(* IEC 61131-3 sources: daoli-st-library/DL_MathData (part 9) *)

(* ---- FC_DL_BcdAddByte.st ---- *)
(*==============================================================================
 * 组件名称 : FC_DL_BcdAddByte ｜ 子库 : DL_MathData ｜ v1.0.0 ｜ 2026-11-23
 * 平台     : CODESYS 3.5 / TwinCAT 3 / InoProShop / Machine Expert（纯 IEC，无厂商库）
 * 功能简介 : 两位 BCD 字节加法：先解码为二进制求和，和 > 99 置错并饱和
 *            到 99，再编码回 BCD。输入含非法 BCD 半字节时置错并返 0。
 * 契约     : 返回 BCD 和 [两位 BCD 形]；xError = TRUE 表示溢出 / 非法输入，
 *            此时返回 99（溢出饱和）或 0（非法输入）；纯函数无状态。
 * 依赖     : 无 DL_ 内部依赖（本批自足实现，不引用库内其他件）
 * 红线自检 : R1 零全局 R2 零%I/%Q R3 纯IEC（*_TO_* 显式转换）
 *            R4 非法 BCD 拒收 + 溢出饱和不回绕 R5 双语注释
 *            R6 N/A（无状态机） R7 N/A（无定时器实例）
 * 修订历史 : 2026-11-23 R78-B1 BCD 校验与算术族模板派生首版
 *============================================================================*)
FUNCTION FC_DL_BcdAddByte : BYTE
VAR_INPUT
    byA : BYTE;         // BCD 加数 / First BCD addend
    byB : BYTE;         // BCD 被加数 / Second BCD addend
END_VAR
VAR_OUTPUT
    xError : BOOL;      // 置错标志：输入非法或和溢出 / Error flag: invalid input or overflow
END_VAR
VAR
    nA : INT;           // byA 解码二进制值 [0..99] / Binary value decoded from byA
    nB : INT;           // byB 解码二进制值 [0..99] / Binary value decoded from byB
    nS : INT;           // 二进制和 [0..99] / Binary sum
    nTens : INT;        // 十位数字 [0..9] / Tens digit
    nOnes : INT;        // 个位数字 [0..9] / Ones digit
END_VAR
xError := FALSE;                    // 置错标志预清 / Preset error flag cleared
FC_DL_BcdAddByte := 16#00;          // 返回值预置 0 / Preset return 0
IF ((byA AND 16#0F) > 16#09) OR (SHR(byA, 4) > 16#09)
    OR ((byB AND 16#0F) > 16#09) OR (SHR(byB, 4) > 16#09) THEN
    xError := TRUE;                 // 输入含非法 BCD 半字节 / Invalid BCD nibble in input
    RETURN;
END_IF
nA := BYTE_TO_INT(SHR(byA, 4)) * 10 + BYTE_TO_INT(byA AND 16#0F);   // 解码 byA / Decode byA
nB := BYTE_TO_INT(SHR(byB, 4)) * 10 + BYTE_TO_INT(byB AND 16#0F);   // 解码 byB / Decode byB
nS := nA + nB;                      // 二进制求和 / Binary sum
IF nS > 99 THEN
    xError := TRUE;                 // 和溢出两位 BCD 域 / Sum overflows two-digit BCD
    nS := 99;                       // 饱和到 99，不回绕 / Saturate at 99, no wrap
END_IF
nTens := nS / 10;                   // 取十位 / Extract tens digit
nOnes := nS MOD 10;                 // 取个位 / Extract ones digit
FC_DL_BcdAddByte := SHL(INT_TO_BYTE(nTens), 4) OR INT_TO_BYTE(nOnes);   // 编码回 BCD / Encode back to BCD
END_FUNCTION

(* ---- FC_DL_BcdDecrementByte.st ---- *)
(*==============================================================================
 * 组件名称 : FC_DL_BcdDecrementByte ｜ 子库 : DL_MathData ｜ v1.0.0 ｜ 2026-11-23
 * 平台     : CODESYS 3.5 / TwinCAT 3 / InoProShop / Machine Expert（纯 IEC，无厂商库）
 * 功能简介 : BCD 字节减 1（如计数值递减）：0 借位回 99（循环计数口径）。
 *            输入含非法 BCD 半字节时防御性返回 0。
 * 契约     : 返回 BCD 减 1 结果 [两位 BCD 形]；非法输入返回 0；
 *            纯函数无状态、同输入同输出。
 * 依赖     : 无 DL_ 内部依赖（本批自足实现，不引用库内其他件）
 * 红线自检 : R1 零全局 R2 零%I/%Q R3 纯IEC（*_TO_* 显式转换）
 *            R4 非法 BCD 返 0 + 0 借位回 99 不越域 R5 双语注释
 *            R6 N/A（无状态机） R7 N/A（无定时器实例）
 * 修订历史 : 2026-11-23 R78-B1 BCD 校验与算术族模板派生首版
 *============================================================================*)
FUNCTION FC_DL_BcdDecrementByte : BYTE
VAR_INPUT
    byVal : BYTE;       // 待递减 BCD 字节 / BCD byte to be decremented
END_VAR
VAR
    nV : INT;           // 解码二进制值 [0..99] / Decoded binary value
    nTens : INT;        // 十位数字 [0..9] / Tens digit
    nOnes : INT;        // 个位数字 [0..9] / Ones digit
END_VAR
FC_DL_BcdDecrementByte := 16#00;    // 返回值预置 0 / Preset return 0
IF ((byVal AND 16#0F) > 16#09) OR (SHR(byVal, 4) > 16#09) THEN
    RETURN;                         // 非法 BCD 输入防御性返 0 / Invalid BCD input returns 0
END_IF
nV := BYTE_TO_INT(SHR(byVal, 4)) * 10 + BYTE_TO_INT(byVal AND 16#0F);   // 解码 / Decode
nV := nV - 1;                       // 二进制减 1 / Decrement in binary
IF nV < 0 THEN
    nV := 99;                       // 0 借位回 99 / Borrow 0 back to 99
END_IF
nTens := nV / 10;                   // 取十位 / Extract tens digit
nOnes := nV MOD 10;                 // 取个位 / Extract ones digit
FC_DL_BcdDecrementByte := SHL(INT_TO_BYTE(nTens), 4) OR INT_TO_BYTE(nOnes);     // 编码回 BCD / Encode back to BCD
END_FUNCTION

(* ---- FC_DL_BcdIncrementByte.st ---- *)
(*==============================================================================
 * 组件名称 : FC_DL_BcdIncrementByte ｜ 子库 : DL_MathData ｜ v1.0.0 ｜ 2026-11-23
 * 平台     : CODESYS 3.5 / TwinCAT 3 / InoProShop / Machine Expert（纯 IEC，无厂商库）
 * 功能简介 : BCD 字节加 1（如计数器 / 计数值递增）：99 进位回 0。
 *            输入含非法 BCD 半字节时防御性返回 0。
 * 契约     : 返回 BCD 加 1 结果 [两位 BCD 形]；非法输入返回 0；
 *            纯函数无状态、同输入同输出。
 * 依赖     : 无 DL_ 内部依赖（本批自足实现，不引用库内其他件）
 * 红线自检 : R1 零全局 R2 零%I/%Q R3 纯IEC（*_TO_* 显式转换）
 *            R4 非法 BCD 返 0 + 99 进位回 0 不越域 R5 双语注释
 *            R6 N/A（无状态机） R7 N/A（无定时器实例）
 * 修订历史 : 2026-11-23 R78-B1 BCD 校验与算术族模板派生首版
 *============================================================================*)
FUNCTION FC_DL_BcdIncrementByte : BYTE
VAR_INPUT
    byVal : BYTE;       // 待递增 BCD 字节 / BCD byte to be incremented
END_VAR
VAR
    nV : INT;           // 解码二进制值 [0..99] / Decoded binary value
    nTens : INT;        // 十位数字 [0..9] / Tens digit
    nOnes : INT;        // 个位数字 [0..9] / Ones digit
END_VAR
FC_DL_BcdIncrementByte := 16#00;    // 返回值预置 0 / Preset return 0
IF ((byVal AND 16#0F) > 16#09) OR (SHR(byVal, 4) > 16#09) THEN
    RETURN;                         // 非法 BCD 输入防御性返 0 / Invalid BCD input returns 0
END_IF
nV := BYTE_TO_INT(SHR(byVal, 4)) * 10 + BYTE_TO_INT(byVal AND 16#0F);   // 解码 / Decode
nV := nV + 1;                       // 二进制加 1 / Increment in binary
IF nV > 99 THEN
    nV := 0;                        // 99 进位回 0 / Carry 99 back to 0
END_IF
nTens := nV / 10;                   // 取十位 / Extract tens digit
nOnes := nV MOD 10;                 // 取个位 / Extract ones digit
FC_DL_BcdIncrementByte := SHL(INT_TO_BYTE(nTens), 4) OR INT_TO_BYTE(nOnes);     // 编码回 BCD / Encode back to BCD
END_FUNCTION

(* ---- FC_DL_BcdIsValidByte.st ---- *)
(*==============================================================================
 * 组件名称 : FC_DL_BcdIsValidByte ｜ 子库 : DL_MathData ｜ v1.0.0 ｜ 2026-11-23
 * 平台     : CODESYS 3.5 / TwinCAT 3 / InoProShop / Machine Expert（纯 IEC，无厂商库）
 * 功能简介 : 判定字节是否为合法两位 BCD 编码：高 / 低半字节均须 <= 9
 *            （0x0A..0x0F 非法）。纯位运算实现，不用库函数。
 * 契约     : 返回 TRUE = 合法 BCD 字节（00..99 的 BCD 形）；输入 byVal
 *            任意字节；纯函数无状态、同输入同输出。
 * 依赖     : 无 DL_ 内部依赖（本批自足实现）
 * 红线自检 : R1 零全局 R2 零%I/%Q R3 纯IEC R4 半字节越 9 拒收
 *            R5 双语注释 R6 N/A（无状态机） R7 N/A（无定时器实例）
 * 修订历史 : 2026-11-23 R78-B1 BCD 校验与算术族模板派生首版
 *============================================================================*)
FUNCTION FC_DL_BcdIsValidByte : BOOL
VAR_INPUT
    byVal : BYTE;       // 待判定字节 / Byte to be validated
END_VAR
IF ((byVal AND 16#0F) > 16#09) OR (SHR(byVal, 4) > 16#09) THEN
    FC_DL_BcdIsValidByte := FALSE;      // 任一半字节 > 9：非法 BCD / Any nibble > 9: invalid BCD
ELSE
    FC_DL_BcdIsValidByte := TRUE;       // 高低半字节均 <= 9：合法 / Both nibbles <= 9: valid
END_IF
END_FUNCTION

(* ---- FC_DL_BcdIsValidWord.st ---- *)
(*==============================================================================
 * 组件名称 : FC_DL_BcdIsValidWord ｜ 子库 : DL_MathData ｜ v1.0.0 ｜ 2026-11-23
 * 平台     : CODESYS 3.5 / TwinCAT 3 / InoProShop / Machine Expert（纯 IEC，无厂商库）
 * 功能简介 : 判定 16 位字是否为合法 4 位 BCD 编码：4 个半字节均须 <= 9
 *            （任一半字节 0x0A..0x0F 非法）。纯位运算 FOR 循环实现，
 *            不用库函数。
 * 契约     : 返回 TRUE = 合法 BCD 字（0000..9999 的 BCD 形）；输入 wVal
 *            任意字；循环轮次固定 4，结构有界；纯函数无状态。
 * 依赖     : 无 DL_ 内部依赖（本批自足实现）
 * 红线自检 : R1 零全局 R2 零%I/%Q R3 纯IEC R4 半字节越 9 拒收 + FOR 上界常量
 *            R5 双语注释 R6 N/A（无状态机） R7 N/A（无定时器实例）
 * 修订历史 : 2026-11-23 R78-B1 BCD 校验与算术族模板派生首版
 *============================================================================*)
FUNCTION FC_DL_BcdIsValidWord : BOOL
VAR_INPUT
    wVal : WORD;        // 待判定 16 位字 / Word to be validated
END_VAR
VAR
    i : INT;            // 半字节序号 0..3 / Nibble index 0..3
END_VAR
FC_DL_BcdIsValidWord := TRUE;       // 预置合法，逐位复核 / Preset valid, recheck nibble by nibble
FOR i := 0 TO 3 DO                  // 4 个半字节逐一校验 / Check all 4 nibbles
    IF (SHR(wVal, i * 4) AND 16#000F) > 16#0009 THEN
        FC_DL_BcdIsValidWord := FALSE;      // 该半字节 > 9：非法 BCD / Nibble > 9: invalid BCD
    END_IF
END_FOR
END_FUNCTION

(* ---- FC_DL_BcdSubByte.st ---- *)
(*==============================================================================
 * 组件名称 : FC_DL_BcdSubByte ｜ 子库 : DL_MathData ｜ v1.0.0 ｜ 2026-11-23
 * 平台     : CODESYS 3.5 / TwinCAT 3 / InoProShop / Machine Expert（纯 IEC，无厂商库）
 * 功能简介 : 两位 BCD 字节减法：先解码为二进制求差，差 < 0（借位下溢）
 *            置错并饱和到 0，再编码回 BCD。输入含非法 BCD 半字节时置错
 *            并返 0。
 * 契约     : 返回 BCD 差 [两位 BCD 形]；xError = TRUE 表示下溢 / 非法输入，
 *            此时返回 0（下溢饱和）；纯函数无状态。
 * 依赖     : 无 DL_ 内部依赖（本批自足实现，不引用库内其他件）
 * 红线自检 : R1 零全局 R2 零%I/%Q R3 纯IEC（*_TO_* 显式转换）
 *            R4 非法 BCD 拒收 + 下溢饱和不回绕 R5 双语注释
 *            R6 N/A（无状态机） R7 N/A（无定时器实例）
 * 修订历史 : 2026-11-23 R78-B1 BCD 校验与算术族模板派生首版
 *============================================================================*)
FUNCTION FC_DL_BcdSubByte : BYTE
VAR_INPUT
    byA : BYTE;         // BCD 被减数 / BCD minuend
    byB : BYTE;         // BCD 减数 / BCD subtrahend
END_VAR
VAR_OUTPUT
    xError : BOOL;      // 置错标志：输入非法或借位下溢 / Error flag: invalid input or borrow underflow
END_VAR
VAR
    nA : INT;           // byA 解码二进制值 [0..99] / Binary value decoded from byA
    nB : INT;           // byB 解码二进制值 [0..99] / Binary value decoded from byB
    nD : INT;           // 二进制差 [0..99] / Binary difference
    nTens : INT;        // 十位数字 [0..9] / Tens digit
    nOnes : INT;        // 个位数字 [0..9] / Ones digit
END_VAR
xError := FALSE;                    // 置错标志预清 / Preset error flag cleared
FC_DL_BcdSubByte := 16#00;          // 返回值预置 0 / Preset return 0
IF ((byA AND 16#0F) > 16#09) OR (SHR(byA, 4) > 16#09)
    OR ((byB AND 16#0F) > 16#09) OR (SHR(byB, 4) > 16#09) THEN
    xError := TRUE;                 // 输入含非法 BCD 半字节 / Invalid BCD nibble in input
    RETURN;
END_IF
nA := BYTE_TO_INT(SHR(byA, 4)) * 10 + BYTE_TO_INT(byA AND 16#0F);   // 解码 byA / Decode byA
nB := BYTE_TO_INT(SHR(byB, 4)) * 10 + BYTE_TO_INT(byB AND 16#0F);   // 解码 byB / Decode byB
nD := nA - nB;                      // 二进制求差 / Binary difference
IF nD < 0 THEN
    xError := TRUE;                 // 借位下溢出两位 BCD 域 / Borrow underflow
    nD := 0;                        // 饱和到 0，不回绕 / Saturate at 0, no wrap
END_IF
nTens := nD / 10;                   // 取十位 / Extract tens digit
nOnes := nD MOD 10;                 // 取个位 / Extract ones digit
FC_DL_BcdSubByte := SHL(INT_TO_BYTE(nTens), 4) OR INT_TO_BYTE(nOnes);   // 编码回 BCD / Encode back to BCD
END_FUNCTION

(* ---- FC_DL_BcdToByte.st ---- *)
(*
    FC_DL_BcdToByte —— 2 位半字节 BCD 解码（BYTE 容器）
    ------------------------------------------------------------------
    分类      : DL_MathData / Convert
    前缀      : FC_DL_
    版本      : 1.0.0
    溯源      : IEC 61131-3 标准语义的道莅防御性实现（BYTE 容器 2 位 BCD → USINT 数值）；
                域内委托平台内建 BCD_TO_BYTE，本件不重实现数学内核；
                半字节合法性校验、满量程提示、错误分级与码位 100% 自有；
                clean-room 重写，未复制任何闭源厂商源码，参考实现仅限 MIT/Apache 许可
    平台      : 纯 IEC 61131-3，CODESYS V3.5+ / TwinCAT 3 / InoProShop 通用
    作者      : 道莅代码库 · PLC编程专家（R20）
    ------------------------------------------------------------------
    功能说明  : 拨码开关组态位、老式仪表组态字最常见的 2 位 BCD 编码（一个 BYTE 装 0~99），
                解码成 0~99 的数值参与比对。
                核心防御：① 先判后算——两个半字节都必须 ≤ 9 才允许进内建。
                   非法 BCD（如 16#1F、16#AA）在内建层的行为平台各不相同（有的翻转、
                   有的返回原值、有的置 0），是本件最不能容忍的不确定点；
                ② 校验只看半字节数值，不看容器大小，故 16#99 合法、16#FF 非法；
                ③ 满量程 99 发信息级提示：拨码全拨到 9 常是调试残留，
                   值本身合法，不该升故障级；
                ④ 合成路径（若平台缺内建）在容器校验之后做半字节乘加，
                   属校验后合成，不是重实现数学内核。
                职责边界：反向编码归 FC_DL_ByteToBcd；4 位 Word 容器归 FC_DL_BcdToWord，
                8 位 Udint 容器归 FC_DL_BcdToUdint；本件只管 2 位拨码容器。
    编译门槛  : 主路径依赖平台内建 BCD_TO_BYTE，三平台标准库均提供。
                若目标平台缺该内建，按合成路径落地：uOut = uHi * 10 + uLo，
                两半字节已由段 2 保证 ≤ 9，乘加结果必然 ≤ 99，无溢出可能。
    错误码    : 16#0001_041C BCD 值恰为满量程 99（多拨码开关调试残留）——信息级，值可用
                16#0001_041D 预留禁用（信息级，不得挪用）
                16#0001_0348 非法 BCD（某半字节 > 9）——故障级，返回 0
                16#0001_0349 预留（故障级，不得挪用）
                16#0001_034A 预留禁用（故障级，不得挪用）
    码位总账  : 16#0001_041C 用 / 16#0001_041D 预留 ｜ 16#0001_0348 用 / 16#0001_0349 预留 / 16#0001_034A 预留
    状态机    : R6 标注 N/A —— 本组件为纯函数无顺序状态机，无 CASE 可写，非法状态不可能出现
    采样约定  : 本件无定时器、无沿检测、无状态；单拍纯计算，结论与任务周期无关。
    修订记录  : 2026-11-16 v1.0.0 首次入库（R20）
*)
FUNCTION FC_DL_BcdToByte : USINT
VAR_INPUT
    uBcd             : BYTE;                  // BCD 编码值 [无量纲]，每半字节 0~9，合计 0~99 / BCD value [dimensionless], each nibble 0 to 9, total 0 to 99
END_VAR
VAR_OUTPUT
    eErr             : UDINT;                 // 错误码，0=正常 / error id, 0=ok
    bError           : BOOL;                  // 故障标志，eErr 为故障级时 TRUE / error flag, TRUE on fault-level eErr
    bValid           : BOOL;                  // 返回值是否可用（非法 BCD 为 FALSE）/ return usable, FALSE on an illegal BCD
END_VAR
VAR CONSTANT
    DL_BCD_NIB_MAX   : BYTE := 9;             // 单个半字节的合法上限 [无量纲] / legal upper bound of one nibble [dimensionless]
    DL_BCD_MASK_LO   : BYTE := 16#0F;         // 低半字节掩码 [位图] / low nibble mask [bitmap]
    DL_BCD_SHIFT_HI  : USINT := 4;            // 高半字节移位量 [bit]，结构性小于 8 / the high nibble shift [bit], structurally below 8
    DL_BCD_FULL      : USINT := 99;           // 满量程值，用于提示 [无量纲] / full scale value used by the hint [dimensionless]
    DL_USINT_ZERO    : USINT := 0;            // 无符号零常量，避免裸字面量 [无量纲] / unsigned zero constant [dimensionless]
END_VAR
VAR
    uLo              : BYTE;                  // 低半字节 [无量纲] / the low nibble [dimensionless]
    uHi              : BYTE;                  // 高半字节 [无量纲] / the high nibble [dimensionless]
    uOut             : USINT;                 // 结果中间量 [无量纲] / result intermediate [dimensionless]
END_VAR

// 段 1｜返回值与错误状态预置 / segment 1, preset return value and error status
FC_DL_BcdToByte := DL_USINT_ZERO;             // 故障缺省返回 0 [无量纲] / fault default returns zero [dimensionless]
eErr := 0;                                    // 预置无错误 / preset no error
bError := FALSE;                              // 预置无故障 / preset no fault
bValid := FALSE;                              // 预置不可用，通过闸门后置位 / preset invalid, set TRUE after the gates
uOut := DL_USINT_ZERO;                        // 结果中间量清零 / clear the result intermediate

// 段 2｜半字节分解与合法性校验（先判后算，域外绝不进内建）/ segment 2, nibble split and legality gate
uLo := uBcd AND DL_BCD_MASK_LO;               // 低半字节 [无量纲] / extract the low nibble [dimensionless]
uHi := SHR(uBcd, DL_BCD_SHIFT_HI);            // 高半字节，移位量 4 结构性小于 8 [无量纲] / extract the high nibble, the shift stays below 8 [dimensionless]

IF (uLo > DL_BCD_NIB_MAX) OR (uHi > DL_BCD_NIB_MAX) THEN
    eErr := 16#0001_0348;                     // 故障级：非法 BCD，半字节超 9 / fault level, illegal BCD, a nibble exceeds nine
    bError := TRUE;                           // 置故障标志 / raise the error flag
    bValid := FALSE;                          // 返回值不可用 / flag the return as unusable
    FC_DL_BcdToByte := DL_USINT_ZERO;         // 确定缺省值 0 / deterministic default of zero
    RETURN;                                   // 出口，不触碰内建 / exit, the built-in is never touched
END_IF

// 段 3｜主体：容器校验通过后委托平台内建 / segment 3, delegate the built-in after the container check
uOut := BYTE_TO_USINT(BCD_TO_BYTE(uBcd));     // BCD → 数值 [无量纲] / decode BCD into a number [dimensionless]

// 段 4｜发布结果与满量程提示（信息级，不置 bError）/ segment 4, publish and hint the full scale value
FC_DL_BcdToByte := uOut;                      // 输出解码值 0~99 [无量纲] / publish the decoded value 0 to 99 [dimensionless]
bValid := TRUE;                               // 合法 BCD 即可用 / a legal BCD is usable
IF uOut = DL_BCD_FULL THEN
    eErr := 16#0001_041C;                     // 信息级：满量程 99，多为拨码调试残留 / info level, full scale, often left over from commissioning
END_IF
END_FUNCTION

(* ---- FC_DL_BcdToDint.st ---- *)
(*
  ==================================================================
  组件名 Component  : FC_DL_BcdToDint
  分类   Category   : DL_MathData
  前缀   Naming     : FC_DL_ ｜ b/n/u/f/t/e/st 类型前缀制（R265）
  码位   Code ID    : 16#0001_0657（故障级）
  版本   Version    : 1.0.0
  复杂度 Complexity  : 低
  功能   Purpose    : 8 位 BCD（DWORD 容器，8 个半字节）→ DINT，逐码元合法性闸，
                      任一半字节 > 9 判故障早退，禁静默按半字节折算。
  开源溯源 Origin    : 公开公式 clean-room，参考 BCD 编码公开工程语义（分类与参数域
                      借鉴，零代码复制），本件实现、闸门与码位 100% 自有。
  许可证 License    : MIT
  参考   Reference  : IEC 61131-3:2013 §6.6 移位与位运算符（SHR / AND）
  平台   Platform   : 纯 IEC 61131-3（FOR / SHR / AND / 四则），三平台通用
  依赖   Depends    : 仅 Standard.library（无库调用）
  分工声明 Split     : FC_DL_BcdToByte / FC_DL_BcdToWord / FC_DL_BcdToUdint 为既有
                      BCD 解码族（BYTE / WORD / UDINT 位宽），本件补 DWORD 8 位宽
                      解码口，四件互引（R216）。
  归属 Ownership     : 本件无 TYPE 声明；全部引脚为 IEC 标准原生类型。
  ------------------------------------------------------------------
  边界 Boundary     :
                      一 域证明（写死）：8 位 BCD 最大 99999999 < 2147483647（DINT
                         上界），累加无溢出可能，故本件无溢出分支；
                      二 逐码元提取：SHR 移位量 4·k（k = 0..7）最大 28 < 32（DWORD
                         位宽），结构性安全（R48 移位量归一：移位量上界由循环界
                         常量证明，禁运行时可变移位量越位宽）；
                      三 任一码元 > 9 → 故障级码 + bBadDigit = TRUE + nOut = 0 +
                         三件套 + RETURN 早退（禁把 A~F 半字节静默折算）；
                      四 首个非法码元即早退（首因保序），bBadDigit 单点置位；
                      五 纯函数：无记忆量、无定时器、无边沿实例，每调用重算；
                      六 无全局、无外部变量、无物理地址、无指针。
  错误码 Codes      :
    16#0001_0657【故障级】非法码元（8 个半字节任一 > 9，首个非法位即早退）
  码位反证 Note     :
    本件仅一个故障场景：8 个码元的合法性出口组合完全同形（nOut = 0、bBadDigit =
    TRUE、bValid = FALSE），无法从输出区分「哪一位非法」，按 R90 只立一码，
    非法位序号不外显（如需位级定位由调用方自行逐半字节复扫）。
  验收 Acceptance   :
    算法已证（脚本）：未跑 ｜ 编译器已证（三平台）：未跑
    V1 16#00000000 → 0；V2 16#99999999 → 99999999（精确无溢出）
    V3 16#0000000A → 故障 0657 + bBadDigit（禁折算）
    V4 16#12345678 → 12345678；V5 16#00000007 → 7（前导零）
    V6 高位半字节 16#A0000000 与低位 16#0000000F → 均故障（A/F 两端抽验）
  修订记录 Revision  :
    2026-11-21  v1.0.0  R63 首版（批 1 · 序号 1）
  ==================================================================
*)
FUNCTION FC_DL_BcdToDint : BOOL
VAR_INPUT
    udBcd   : DWORD := 16#00000000; // 8 位 BCD 输入 [码]，8 个半字节 / the eight digit BCD input in a double word container
END_VAR
VAR_OUTPUT
    nOut    : DINT := 0;            // 解码结果 [个]，非法码元时为 0 / the decoded result, zero when a digit is illegal
    bBadDigit : BOOL := FALSE;      // 非法码元标志（任一半字节 > 9）[-] / the illegal digit flag raised when any nibble exceeds nine
    bValid  : BOOL := FALSE;        // 结果可用 [-] / the result usable flag
    eErr    : UDINT := 16#0000_0000; // 错误码，0 = 正常 / the error code, zero is ok
    bError  : BOOL := FALSE;        // 故障标志（故障级码同拍置位，R45 配对）/ the fault flag raised with a fault level code
END_VAR
VAR
    k       : DINT := 0;  // 半字节遍历索引 [下标]，0..7 / the nibble traversal index from zero to seven
    nShift  : DINT := 0;  // 移位量 [位]，4·k ≤ 28 结构性安全 / the shift amount of four times the index, proven below the word width
    uDig    : USINT := 0; // 当前半字节码元 [位] / the current digit nibble
    nAcc    : DINT := 0;  // 十进制累加器（Horner 展开）[个] / the decimal accumulator of the Horner expansion
END_VAR  // R64 结构补齐：VAR 段缺失的 END_VAR（门禁机械修复）
VAR CONSTANT
    DL_BCD_MASK  : DWORD := 16#0000000F; // 半字节掩码常量（提级禁魔法数）[-] / the nibble mask constant lifted out of the body
    DL_BCD_DIG9  : USINT := 9;           // 合法码元上界 [位] / the legal digit ceiling of nine
    DL_BCD_NIB   : DINT := 4;            // 每码元位宽 [位] / the nibble width of four bits
    DL_BCD_N     : DINT := 8;            // 码元总数 [个]（DWORD 恰 8 半字节，R57）/ the nibble count of eight aligned with the container
    DL_BCD_ZERO  : DINT := 0;            // 整型零常量 [个] / the integer zero constant
    DL_BCD_ONE   : DINT := 1;            // 整型一常量 [个] / the integer one constant
    DL_BCD_TEN   : DINT := 10;           // 十进制权值基数 [个] / the decimal weight base of ten
END_VAR

// 段 1｜返回值与全部出口预置安全值（R45 四段式第一段）/ segment 1, the preset of the return and every outlet
FC_DL_BcdToDint := FALSE; // 返回值预置假 / preset the return false
nOut := DL_BCD_ZERO; // 结果预置零 [个] / preset the result zero
bBadDigit := FALSE; // 非法码元标志预置假 / preset the illegal digit flag false
bValid := FALSE; // 可用标志预置假 / preset the validity false
eErr := 16#0000_0000; // 错误码预置正常 / preset the code to ok
bError := FALSE; // 故障标志预置假 / preset the error flag false
nAcc := DL_BCD_ZERO; // 累加器预置零 [个] / preset the accumulator zero
k := DL_BCD_ZERO; // 索引预置零 / preset the index zero
nShift := DL_BCD_ZERO; // 移位量预置零 [位] / preset the shift amount zero
uDig := 0; // 码元预置零 [位] / preset the digit zero

// 段 2｜逐码元提取与合法性闸（移位量 4·k ≤ 28 < 32 结构性安全，边界二）/ segment 2, the digit extraction with the structural shift bound
FOR k := DL_BCD_ZERO TO DL_BCD_N - DL_BCD_ONE DO // 有界遍历 8 个半字节（循环界常量证明，无死循环）/ the bounded traversal over eight nibbles proven by the constant loop bound
    nShift := DL_BCD_NIB * k; // 移位量 = 4·k，最大 28 [位] / the shift amount of four times the index, at most twenty eight
    uDig := DWORD_TO_USINT(SHR(udBcd, nShift) AND DL_BCD_MASK); // 提取当前半字节（SHR 后与掩码，常量提级）/ extract the current nibble by shifting then masking with the lifted constant
    IF uDig > DL_BCD_DIG9 THEN // 码元 > 9：非法（边界三，禁折算）/ a digit above nine is illegal, never folded silently
        bBadDigit := TRUE; // 置非法码元标志 / raise the illegal digit flag
        eErr := 16#0001_0657; // 故障级：非法码元 / fault grade, an illegal digit
        bError := TRUE; // 同拍置故障标志（R45 配对）/ raise the fault flag on the same scan
        bValid := FALSE; // 结果不可用 / the result is not usable
        nOut := DL_BCD_ZERO; // 结果强制归零（禁部分折算值外泄）/ force the result to zero so no partial fold leaks
        RETURN; // 早退（首因保序，边界四）/ early return with the first cause kept
    END_IF
    nAcc := (nAcc * DL_BCD_TEN) + USINT_TO_DINT(uDig); // Horner 十进制累加：nAcc = nAcc×10 + 码元 [个] / the Horner decimal accumulation, the domain proof in boundary one covers every step
END_FOR

// 段 3｜统一出口（域证明：nAcc ≤ 99999999 < DINT 上界，无溢出分支，边界一）/ segment 3, the unified outlet with the domain proof
nOut := nAcc; // 结果出口 [个] / the result outlet
bValid := TRUE; // 结果可用 / the result is usable
FC_DL_BcdToDint := TRUE; // 返回成功 / return success
END_FUNCTION

(* ---- FC_DL_BcdToUdint.st ---- *)
(*
    FC_DL_BcdToUdint —— 8 位十进制 BCD 码到 UDINT 防御转换
    ------------------------------------------------------------------
    分类      : DL_MathData / Convert
    前缀      : FC_DL_
    版本      : 1.0.0
    溯源      : IEC 61131-3 标准语义的道莅防御性实现
                （内部委托平台内建函数，外围统一错误码/钳位/双语文档；
                  未复制任何闭源厂商源码，参考实现仅限 MIT/Apache 许可）
    平台      : 纯 IEC 61131-3，CODESYS / TwinCAT / InoProShop 通用
    作者      : 道莅代码库 · PLC编程专家（R16）
    ------------------------------------------------------------------
    功能说明  : 将 8 位十进制 BCD 码输入（每半字节 0~9）防御性转换为 UDINT 并返回；
                逐半字节合法性校验：任一半字节值 > 9（即 16#A~16#F 非法 BCD 码）判为
                故障级 16#0001_02A6，返回 0 且 bValid=FALSE；
                域内按半字节以 10 为基加权累加还原十进制值（乘子为常量基 10 的幂，
                最大权值 10^7、最大累加和 99999999，均在 UDINT 域内无溢出）；
                校验覆盖范围说明：UDINT 为 32 位容器，恰含 8 个 BCD 半字节（k=0..7），
                完整覆盖 8 位十进制域 0..99999999；k=8..15 的半字节在 32 位容器中不存在，
                且移位量 ≥32 属跨平台未定义行为，故不实施越界校验；
                本组件无钳位路径（非法半字节直接故障拦截，域内值精确还原）。
    错误码    : 16#0001_02A6 存在非法 BCD 半字节（半字节值 16#A~16#F）——故障级，返回 0
                16#0001_01D0 预留禁用（信息级，不得挪用）
                16#0001_01D1 预留禁用（信息级，不得挪用）
                16#0001_02A7 预留禁用（故障级，不得挪用）
                16#0001_02A8 预留禁用（故障级，不得挪用）
    状态机    : R6 标注 N/A —— 本组件为纯函数无顺序状态机，无 CASE 可写，非法状态不可能出现，故以本节说明替代 ELSE 兜底
    修订记录  : 2026-11-16 v1.0.0 首次入库（R16）
*)
FUNCTION FC_DL_BcdToUdint : UDINT
VAR_INPUT
    uBcd : UDINT; // 8 位十进制 BCD 码 [BCD 位]，每半字节 0~9 / 8-digit BCD code, each nibble 0~9
END_VAR
VAR_OUTPUT
    eErr   : UDINT; // 错误码，0=正常 / error id, 0=ok
    bError : BOOL;  // 是否出错，eErr 非 0 时为 TRUE / error flag, TRUE when eErr is nonzero
    bValid : BOOL;  // 输出是否有效可用 / output valid flag
END_VAR
VAR CONSTANT
    DL_BCD_NIB_MASK : UDINT := 16#F;  // 半字节掩码 [BCD 位] / nibble mask
    DL_BCD_NIB_MAX  : UDINT := 16#9;  // 合法 BCD 半字节上界 9 [BCD 位] / valid BCD nibble upper bound 9
    DL_BCD_NIB_CNT  : INT   := 8;     // UDINT 32 位容器 BCD 半字节总数 [个] / total BCD nibble count of 32-bit UDINT container
    DL_DEC_BASE     : UDINT := 10;    // 十进制加权基 [基数] / decimal weighting base
END_VAR
VAR
    i       : INT;   // 半字节循环索引 [个] / nibble loop index
    uNib    : UDINT; // 当前半字节值 [BCD 位] / current nibble value
    uWeight : UDINT; // 当前半字节十进制权值（10^i） [倍] / current nibble decimal weight (10^i)
END_VAR

// 段 1｜返回值与错误状态预置 / segment 1, preset return value and error status
FC_DL_BcdToUdint := 0; // 故障缺省返回 0 [无量纲] / fault default returns 0
eErr   := 0;     // 预置无错误 / preset no error
bError := FALSE; // 预置无故障 / preset no fault
bValid := FALSE; // 预置无效，通过全半字节校验后置位 / preset invalid, set TRUE after all-nibble check passes

// 段 2｜逐半字节校验与十进制加权累加（末段） / segment 2, per-nibble validation and decimal weighted accumulation (final)
uWeight := 1; // 最低半字节权值 10^0 [倍] / lowest nibble weight 10^0
FOR i := 0 TO DL_BCD_NIB_CNT - 1 DO
    uNib := SHR(uBcd, 4 * i) AND DL_BCD_NIB_MASK; // 取第 i 个半字节（SHR 移位量 4*i ≤ 28 安全） / extract i-th nibble (shift 4*i <= 28, safe)
    IF uNib > DL_BCD_NIB_MAX THEN
        FC_DL_BcdToUdint := 0;    // 故障级返回 0，清除部分累加值 / fault level returns 0, clear partial accumulation
        eErr   := 16#0001_02A6;   // 非法 BCD 半字节故障码 / invalid BCD nibble fault id
        bError := TRUE;           // 置故障标志 / set fault flag
        bValid := FALSE;          // 输出无效 / output invalid
        RETURN;                   // 立即返回 / immediate return
    END_IF
    FC_DL_BcdToUdint := FC_DL_BcdToUdint + uNib * uWeight; // 半字节加权累加（最大 99999999 无溢出） / weighted accumulation (max 99999999, no overflow)
    uWeight := uWeight * DL_DEC_BASE; // 权值升位 ×10（最大 10^7，UDINT 域内无溢出） / weight times 10 (max 10^7, no UDINT overflow)
END_FOR
bError := FALSE; // 全部半字节合法，无故障 / all nibbles valid, no fault
bValid := TRUE;  // 输出有效可用 / output valid
END_FUNCTION

(* ---- FC_DL_BilinearInterp.st ---- *)
(*
  ==================================================================
  组件名 Component  : FC_DL_BilinearInterp
  分类   Category   : DL_MathData
  版本   Version    : 1.0.0
  功能   Purpose    : 双线性插值：在等距网格表上按 (fX, fY) 求插值。
                      越界策略=「钳位到边界单元并置码不静默」（头注定稿口径）：
                      fX/fY 超出 [fX0, fX0+(n-1)*d] 时钳到边界单元继续插值，
                      输出有效但带码 02；末端格点用 1E-9 容差处理防 i1 越界
                      一行（fU 恰好等于上界时 i0 退到 n-2、tx 收满 1.0，
                      n=1 退化为常量直通）。
  来源   Source     : t2-1-lgf-math（数学族：双线性插值为公开数值方法口径，
                      实现零源码复制）
  互引   Cross-ref  : FC_DL_InterpolateTable3D（同族三维插值原子，本件为其
                      二维退化对偶，可级联使用）
  平台   Platform   : 纯 IEC 61131-3 四则 + TRUNC，三平台通用
  依赖   Depends    : 无 DL_ 内部依赖；无标准库
  表格口径 Table    : aTable 为定长容量数组（NY_MAX × NX_MAX 见常量段），
                      实际使用 ny=nRows / nx=nCols 由输入给定，容量外元素
                      永不访问（下标闸先行）；行序 = [y 索引][x 索引]。
  红线   Redline    : R1 零全局/VAR_EXTERNAL/R2 零 %I/%Q/R3 纯 IEC 标准
                      R4 步距≤0 与行列数<1 配置闸 + 元素级非有限闸（含四角
                      值）+ 越界钳位显式置码 + 除法分母已闸
                      R5 全变量双语同行注释/R6 纯函数无状态机（CASE 不适用）
                      R7 无定时器与沿检测/R8 容差与容量常量化
  错误码 Codes      : 01【失效级】配置非法（nRows/nCols < 1 或步距 ≤ 0 或
                      行列数超容量），返回 0
                      02【信息级】fX/fY 越界已钳位到边界单元（输出有效）
                      03【失效级】任一输入或四角表值非有限，返回 0
  码位反证 Note     : 02 与 03 分立依据（R90）：02 时 bValid=TRUE 带码、
                      03 时 bValid=FALSE，双通道可唯一区分；01 与 03 分立：
                      01 在配置面可观测、03 在数据面可观测，入口不同。
  验收   Acceptance : V1 网格中心点 → 精确双线性值 ｜ V2 fX 超上界 → 钳边界
                      + 码 02 ｜ V3 fDx=0 → 码 01 ｜ V4 nCols=1 → y 向插值
                      常量直通 ｜ V5 表值 NaN → 码 03 ｜ V6 末端格点容差 →
                      不越界不置 02
  变更   Revision   : 2026-11-22  v1.0.0  R66 首版（编码阶段批 2 序 5）
  ==================================================================
*)
FUNCTION FC_DL_BilinearInterp : LREAL
VAR_INPUT
    aTable : ARRAY[0..BIL_NY_MAX - 1, 0..BIL_NX_MAX - 1] OF LREAL; // 容量网格表 [表值]（实际 ny/nx 由 nRows/nCols 给定，行序=[y][x]）/ the capacity grid table
    nRows  : UDINT;  // 实际行数（y 向格点数）[个]，≥1 / the actual rows, at least one
    nCols  : UDINT;  // 实际列数（x 向格点数）[个]，≥1 / the actual columns, at least one
    fX     : LREAL;  // 查询点 x 坐标 [物理单位同表] / the query x coordinate
    fY     : LREAL;  // 查询点 y 坐标 [物理单位同表] / the query y coordinate
    fX0    : LREAL;  // x 起始格点坐标 [物理单位同表] / the x grid origin
    fDx    : LREAL;  // x 步距 [物理单位同表]，须 > 0 / the x step, must be positive
    fY0    : LREAL;  // y 起始格点坐标 [物理单位同表] / the y grid origin
    fDy    : LREAL;  // y 步距 [物理单位同表]，须 > 0 / the y step, must be positive
END_VAR
VAR_OUTPUT
    bValid : BOOL;   // 输出可用标志（码 02 时仍 TRUE）[-] / the output usable flag, true also with code 02
    nErrId : UDINT;  // 错误码，0=正常，01/02/03 见头注 [码] / the error code [code]
END_VAR
VAR
    fU     : LREAL;  // x 向规格化浮点下标 [格] / the normalized floating x index [cell]
    fV     : LREAL;  // y 向规格化浮点下标 [格] / the normalized floating y index [cell]
    fXmax  : LREAL;  // x 上边界格点坐标 [物理单位] / the x upper boundary coordinate
    fYmax  : LREAL;  // y 上边界格点坐标 [物理单位] / the y upper boundary coordinate
    ix0    : UDINT;  // x 向左格点下标 [格] / the left x cell index
    ix1    : UDINT;  // x 向右格点下标 [格] / the right x cell index
    iy0    : UDINT;  // y 向下格点下标 [格] / the lower y cell index
    iy1    : UDINT;  // y 向上格点下标 [格] / the upper y cell index
    fTx    : LREAL;  // x 向格内分数 0~1 [-] / the in cell x fraction
    fTy    : LREAL;  // y 向格内分数 0~1 [-] / the in cell y fraction
    v00    : LREAL;  // 左下角值 [表值] / the lower left corner value
    v10    : LREAL;  // 右下角值 [表值] / the lower right corner value
    v01    : LREAL;  // 左上角值 [表值] / the upper left corner value
    v11    : LREAL;  // 右上角值 [表值] / the upper right corner value
    fRes   : LREAL;  // 插值结果工作寄存器 [表值] / the interpolation working register
END_VAR
VAR CONSTANT
    BIL_NY_MAX   : UDINT := 32;               // 容量行数上限 [行]（头注表格口径）/ the capacity row limit
    BIL_NX_MAX   : UDINT := 32;               // 容量列数上限 [列]（头注表格口径）/ the capacity column limit
    BIL_EPS      : LREAL := 1.0E-9;           // 末端格点容差 [格] / the end cell tolerance [cell]
    BIL_FIN_MAX  : LREAL := 1.7976931348623157E308; // LREAL 有限上限 [无量纲] / the finite LREAL limit
    BIL_ERR_NONE : UDINT := 16#0000_0000;     // 无错误 [码] / no error [code]
    BIL_ERR_CFG  : UDINT := 16#0000_0001;     // 码 01：配置非法 / code 01, illegal configuration
    BIL_ERR_CLAMP: UDINT := 16#0000_0002;     // 码 02：越界钳位（信息级）/ code 02, clamped, info level
    BIL_ERR_NAN  : UDINT := 16#0000_0003;     // 码 03：非有限 / code 03, non finite
END_VAR

// 段 1｜返回值与输出预置 / segment 1, preset the return and outputs
FC_DL_BilinearInterp := 0.0;  // 失效缺省返回 0 / fault default returns zero
bValid := FALSE;              // 预置不可用 / preset unusable
nErrId := BIL_ERR_NONE;       // 预置无错误 / preset no error

// 段 2｜配置闸（码 01，结构 RETURN 早退）：行列数 ≥1 且不超容量 + 双步距 > 0
//      segment 2, the configuration gate, dimensions inside capacity and positive steps
IF (nRows < UDINT#1) OR (nCols < UDINT#1) OR (nRows > BIL_NY_MAX) OR (nCols > BIL_NX_MAX)
   OR (fDx <= 0.0) OR (fDy <= 0.0) THEN
    nErrId := BIL_ERR_CFG;
    RETURN;
END_IF

// 段 3｜标量输入非有限闸（码 03）：查询点/原点/步距全套（R272 闸参数全覆盖）
//      segment 3, the scalar finiteness gate over every floating input
IF (fX <> fX) OR (fY <> fY) OR (fX0 <> fX0) OR (fY0 <> fY0)
   OR (ABS(fX) > BIL_FIN_MAX) OR (ABS(fY) > BIL_FIN_MAX)
   OR (ABS(fX0) > BIL_FIN_MAX) OR (ABS(fY0) > BIL_FIN_MAX) THEN
    nErrId := BIL_ERR_NAN;
    RETURN;
END_IF

// 段 4｜越界钳位：先算边界坐标再钳查询点，钳位即置码 02 不静默
//      segment 4, the range clamp with the explicit code, never silent
fXmax := fX0 + DINT_TO_LREAL(UDINT_TO_DINT(nCols) - 1) * fDx;   // x 上边界坐标 / the x upper boundary
fYmax := fY0 + DINT_TO_LREAL(UDINT_TO_DINT(nRows) - 1) * fDy;   // y 上边界坐标 / the y upper boundary
IF (fX < fX0) OR (fX > fXmax) OR (fY < fY0) OR (fY > fYmax) THEN
    nErrId := BIL_ERR_CLAMP;                                    // 码 02（信息级，bValid 仍 TRUE）/ code 02, still valid
END_IF
IF fX < fX0 THEN fX := fX0; END_IF                              // x 下钳 / clamp x low
IF fX > fXmax THEN fX := fXmax; END_IF                          // x 上钳 / clamp x high
IF fY < fY0 THEN fY := fY0; END_IF                              // y 下钳 / clamp y low
IF fY > fYmax THEN fY := fYmax; END_IF                          // y 上钳 / clamp y high

// 段 5｜规格化浮点下标：分母步距已闸 > 0 / segment 5, normalized indices, steps gated positive
fU := (fX - fX0) / fDx;                                         // x 浮点下标 [格] / the floating x index
fV := (fY - fY0) / fDy;                                         // y 浮点下标 [格] / the floating y index

// 段 6｜末端格点容差处理（防 i1 越界一行）+ n=1 退化闸，二者合一避免 UDINT 回绕：
//      fU 恰为上界时左格点退到 n-2、分数收满 1.0；n=1 时下标收 0、分数归零
//      segment 6, the end cell tolerance and the single cell degeneration, merged so no UDINT wraparound occurs
ix0 := DINT_TO_UDINT(LREAL_TO_DINT(TRUNC(fU)));                 // 截断得左格点（标准转换链）/ truncate to the left cell, standard conversion chain
iy0 := DINT_TO_UDINT(LREAL_TO_DINT(TRUNC(fV)));                // 截断得下格点 / truncate to the lower cell
IF nCols = UDINT#1 THEN                                         // 单列退化：常量直通 / the single column degeneration
    ix0 := UDINT#0;                                             // 下标收 0 / the index to zero
    fTx := 0.0;                                                 // 分数归零 → 只用左值 / the fraction to zero
ELSIF ix0 >= nCols - UDINT#1 THEN                               // 落在末端格点（含 1E-9 抖动）/ landed on the last cell
    ix0 := nCols - UDINT#2;                                     // 退到倒数第二格（n≥2 时安全）/ step back one cell, safe for n at least two
    fTx := 1.0;                                                 // 分数收满 = 右格点值 / full fraction picks the right value
ELSE
    fTx := fU - DINT_TO_LREAL(UDINT_TO_DINT(ix0));              // 格内分数 / the in cell fraction
END_IF
IF nRows = UDINT#1 THEN                                         // 单行退化 / the single row degeneration
    iy0 := UDINT#0;
    fTy := 0.0;
ELSIF iy0 >= nRows - UDINT#1 THEN
    iy0 := nRows - UDINT#2;
    fTy := 1.0;
ELSE
    fTy := fV - DINT_TO_LREAL(UDINT_TO_DINT(iy0));
END_IF

// 段 7｜右/上格点下标（段 6 已保证 ix0 ≤ nCols-2 或 ix0=0 且 nCols=1，ix1 恒 < nCols）
//      segment 7, the right and upper indices, proven inside the table by segment 6
IF ix0 >= nCols - UDINT#1 THEN                                  // 兜底（结构性不可达，留档）/ defensive, unreachable by construction
    ix1 := ix0;                                                 // 收敛为同格 / collapse to the same cell
ELSE
    ix1 := ix0 + UDINT#1;                                       // 正常右格点 / the normal right cell
END_IF
IF iy0 >= nRows - UDINT#1 THEN
    iy1 := iy0;
ELSE
    iy1 := iy0 + UDINT#1;
END_IF

// 段 8｜四角表值非有限闸（码 03）：下标闸已在段 6/7 完成（ix1<nCols，iy1<nRows）
//      segment 8, the four corner finiteness gate, index gates already proven
v00 := aTable[iy0, ix0];                                        // 左下角 / the lower left corner
v10 := aTable[iy0, ix1];                                        // 右下角 / the lower right corner
v01 := aTable[iy1, ix0];                                        // 左上角 / the upper left corner
v11 := aTable[iy1, ix1];                                        // 右上角 / the upper right corner
IF (v00 <> v00) OR (v10 <> v10) OR (v01 <> v01) OR (v11 <> v11)
   OR (ABS(v00) > BIL_FIN_MAX) OR (ABS(v10) > BIL_FIN_MAX)
   OR (ABS(v01) > BIL_FIN_MAX) OR (ABS(v11) > BIL_FIN_MAX) THEN
    nErrId := BIL_ERR_NAN;
    RETURN;
END_IF

// 段 9｜双线性合成（先 x 后 y，分数均在 [0,1] 域内，凸组合有界）
//      segment 9, the bilinear blend, all fractions inside zero to one
fRes := (1.0 - fTx) * v00 + fTx * v10;                          // y0 行内插 [表值] / the lower row blend
fRes := fRes * (1.0 - fTy) + ((1.0 - fTx) * v01 + fTx * v11) * fTy;  // 行间加权 / the row to row blend

// 段 10｜出口 / segment 10, exit
FC_DL_BilinearInterp := fRes;                                   // 发布插值结果 / publish the result
bValid := TRUE;                                                 // 结果可用（含码 02 场景）/ the result is usable, also with code 02
END_FUNCTION

(* ---- FC_DL_BitArrayReverse.st ---- *)
(*==============================================================================
 * 组件名称 (Component)  : FC_DL_BitArrayReverse
 * 所属子库 (Sublibrary) : DL_MathData
 * 归属目录 (Directory)  : C:\Library\DL_MathData
 * 当前版本 (Version)    : 1.0.0
 * 分类/来源标签         : 函数（FUNCTION）· 纯函数 · 位数组段镜像反转
 *                         iec-std-wrapper / bitstring / bit-array
 * 兼容性   (Platform)   : CODESYS 3.5 / TwinCAT 3 / 汇川 InoProShop / 施耐德
 *                         Machine Expert；零库函数依赖，纯标准布尔交换
 * 溯源声明 (Provenance) : IEC 61131-3 标准语义的道莅防御性实现——内部委托平台标准库语义，
 *                         外围统一错误码 / 钳位 / 双语注释，严禁重实现数学内核。
 * 功能一句话 (Summary)  : 位数组指定段的镜像反转（首尾对调向中推进），段域
 *                         双闸（起始下标、段长），空段或单元素恒等返回。
 *
 * 功能描述 (Function)   : 先过段域双闸：起始下标在 0..127 且段长非负且
 *                         起始加段长不越 128 上界，域外拒绝且不触碰数组；
 *                         合法路径用 VAR_IN_OUT 就地交换，双指针向中推进，
 *                         段长小于等于 1 时恒等返回并告知。
 * 与既有件边界 (Boundary): BitArray 族 Extract/Insert/Rotate/SegCopy 覆盖
 *                         取段、插段、循环移位与段复制；本件补镜像反转原子，
 *                         服务 LSB/MSB 序数组整体换序与测试向量构造。
 * 码位说明 (Codes)      : 信息 16#0002_3054 段长小于等于 1，恒等返回
 *                         故障 16#0002_3055 起始下标域外（小于 0 或越上界）
 *                         故障 16#0002_3056 段长域外（负值或越出数组上界）
 *                         段 16#02_3_54~57 首槽信息级、次槽起故障级。
 * 依赖说明 (Depends)    : 无 DL_ 内部依赖；零库函数依赖。
 * 红线自检 (Redline)    : 零全局依赖 ｜ 零 VAR_EXTERNAL ｜ 零 %I/%Q ｜ 纯 IEC 标准库
 *                         循环上界由已闸段参数给定，无越局面
 *                         全变量双语同行注释 ｜ 无定时器实例 ｜ 无状态机
 * 修订历史 (Revision)   : 2026-11-18  v1.0.0  首版入库（R32 · 批 3）
 *============================================================================*)

FUNCTION FC_DL_BitArrayReverse : BOOL
VAR_INPUT
    iStart : INT;                       // 段起始下标 [索引]，域 0 到 127 / Segment start index, 0 to 127
    iLen   : INT;                       // 段长 [位]，域 0 到 128 减起始 / Segment length in bits
END_VAR
VAR_IN_OUT
    aBits  : ARRAY[0..127] OF BOOL;     // 位数组 [位]，就地反转不复制 / Bit array reversed in place
END_VAR
VAR_OUTPUT
    nSwapped : INT;                     // 交换对数 [对]，段长一半向下取整 / Swap pairs, half the length
    uErrorId : UDINT;                   // 事件码，0 表示无事件 / Event code, zero means none
END_VAR
VAR
    bTmp  : BOOL;   // 交换暂存位 [位] / Swap staging bit
    nLo   : INT;    // 左指针 [索引] / Left pointer
    nHi   : INT;    // 右指针 [索引] / Right pointer
    uCode : UDINT;  // 码位暂存，出口单点写入 [码] / Code staging
END_VAR
VAR CONSTANT
    DL_BAR_SIZE : INT := 128;           // 数组位容量 [位]，与声明一致 / Array capacity, matches the declaration
END_VAR

(* 段 1｜输出预置 / Pre-set *)
FC_DL_BitArrayReverse := FALSE;
nSwapped := 0;
uErrorId := 16#0000_0000;
uCode    := 16#0000_0000;

(* 段 2｜起始下标闸：域外拒绝且不触碰数组 / Start index gate: refuse without touching the array *)
IF (iStart < 0) OR (iStart >= DL_BAR_SIZE) THEN
    uErrorId := 16#0002_3055;    // 故障级：起始下标域外 / Fault: start index out of domain
    RETURN;
END_IF

(* 段 3｜段长闸：非负且段尾不越数组上界 / Length gate: non-negative and the tail inside bounds *)
IF (iLen < 0) OR ((iStart + iLen) > DL_BAR_SIZE) THEN
    uErrorId := 16#0002_3056;    // 故障级：段长域外 / Fault: length out of domain
    RETURN;
END_IF

(* 段 4｜恒等早退：空段或单元素无需交换 / Identity exit: nothing to swap *)
IF iLen <= 1 THEN
    uErrorId := 16#0002_3054;    // 信息级：恒等返回 / Info: identity return
    FC_DL_BitArrayReverse := TRUE;
    RETURN;
END_IF

(* 段 5｜双指针镜像交换：向中推进，交会即停 / Two-pointer mirror swap, stop at the meeting point *)
nLo := iStart;                   // 左指针从段首 / Left pointer at the head
nHi := iStart + iLen - 1;        // 右指针从段尾 / Right pointer at the tail
WHILE nLo < nHi DO
    bTmp        := aBits[nLo];   // 暂存左位 / Stage the left bit
    aBits[nLo]  := aBits[nHi];   // 左位取右位 / Left takes the right
    aBits[nHi]  := bTmp;         // 右位取暂存 / Right takes the staged
    nLo := nLo + 1;              // 左推进 / Advance left
    nHi := nHi - 1;              // 右回退 / Retreat right
    nSwapped := nSwapped + 1;    // 交换对计数 / Count the pair
END_WHILE

(* 段 6｜出口：码位单点写入 / Exit: single write point *)
uErrorId := uCode;               // 无事件，保持零 / No event, stays zero
FC_DL_BitArrayReverse := TRUE;
END_FUNCTION

(* ---- FC_DL_BytesToHexString.st ---- *)
(*==============================================================================
 * 组件名称 (Component)  : FC_DL_BytesToHexString
 * 所属子库 (Sublibrary) : DL_MathData
 * 归属目录 (Directory)  : C:\Library\DL_MathData
 * 当前版本 (Version)    : 1.0.0
 * 分类/来源标签         : 函数（FUNCTION）· 纯函数 · 字节数组十六进制编码
 *                         iec-std-wrapper / string / bitstring
 * 兼容性   (Platform)   : CODESYS 3.5 / TwinCAT 3 / 汇川 InoProShop / 施耐德
 *                         Machine Expert；仅用 Standard.library 的 LEN / MID / CONCAT
 * 溯源声明 (Provenance) : IEC 61131-3 标准语义的道莅防御性实现——内部委托平台标准库语义，
 *                         外围统一错误码 / 钳位 / 双语注释，严禁重实现数学内核。
 * 功能一句话 (Summary)  : 字节数组编码为定宽大写十六进制串，每字节恒出两字符，
 *                         空数组返回空串，计数域外与写出异常双重防御。
 *
 * 功能描述 (Function)   : 先做计数域闸（0 到 127），再逐字节拆高低半字节，
 *                         经 '0123456789ABCDEF' 码表定位拼出两字符，出口校验
 *                         写出长度恰为两倍计数；与 DwordToHexString 互补，
 *                         覆盖变长缓冲的报文与日志场景。
 * 与既有件边界 (Boundary): FC_DL_HexStringToLword 为反向解析单字；本件面向
 *                         数组整体编码，不做前缀、不做分隔符、不做小写。
 * 码位说明 (Codes)      : 信息 16#0002_303C 空数组恒等返回（结果空串）
 *                         故障 16#0002_303D 计数域外（小于 0 或大于 127）
 *                         故障 16#0002_303E 写出长度与两倍计数不一致（防御校验）
 *                         段 16#02_3_3C~3F 首槽信息级、次槽起故障级。
 * 依赖说明 (Depends)    : 无 DL_ 内部依赖；仅 Standard.library 的 LEN / MID / CONCAT。
 * 红线自检 (Redline)    : 零全局依赖 ｜ 零 VAR_EXTERNAL ｜ 零 %I/%Q ｜ 纯 IEC 标准库
 *                         无除法故无除零面 ｜ 移位量 4 与 8 恒小于位宽（归一达标）
 *                         全变量双语同行注释 ｜ 无定时器实例
 * 修订历史 (Revision)   : 2026-11-18  v1.0.0  首版入库（R32 · 批 1）
 *============================================================================*)

FUNCTION FC_DL_BytesToHexString : BOOL
VAR_INPUT
    aBytes  : ARRAY[0..127] OF BYTE;    // 源字节数组 [字节]，最多 127 字节 / Source byte array, at most 127 bytes
    nCount  : INT;                      // 参与编码的字节个数 [字节]，域 0 到 127 / Number of bytes to encode, 0 to 127
END_VAR
VAR_OUTPUT
    sHex     : STRING(255);             // 大写十六进制结果 [ASCII]，长度恰为两倍计数 / Uppercase hex result, twice the count
    nWritten : INT;                     // 写出字符数 [字符] / Characters written
    uErrorId : UDINT;                   // 事件码，0 表示无事件 / Event code, zero means none
END_VAR
VAR
    sTmp   : STRING(255); // 结果累积缓冲 [ASCII] / Result staging buffer
    bCur   : BYTE;        // 当前字节 [字节] / Current byte
    nHi    : INT;         // 高半字节码表下标 [索引] / High nibble table index
    nLo    : INT;         // 低半字节码表下标 [索引] / Low nibble table index
    nI     : INT;         // 字节循环下标 [索引] / Byte loop index
    uCode  : UDINT;       // 码位暂存，出口单点写入 [码] / Code staging
END_VAR
VAR CONSTANT
    DL_BTH_MAXN : INT := 127;               // 最大字节数 [字节]，两倍后仍在 255 内 / Max bytes, doubled stays within 255
    DL_BTH_ONE  : INT := 1;                 // 单字符长度参数 [字符] / Single character length argument
END_VAR

(* 段 1｜输出预置与残留清除 / Pre-set and clear before any branch *)
FC_DL_BytesToHexString := FALSE;
sHex     := '';
sTmp     := '';
nWritten := 0;
uErrorId := 16#0000_0000;
uCode    := 16#0000_0000;

(* 段 2｜计数域闸：契约参数不钳位，域外直接拒绝 / Count gate: a contract value is never clamped *)
IF (nCount < 0) OR (nCount > DL_BTH_MAXN) THEN
    uErrorId := 16#0002_303D;    // 故障级：计数域外 / Fault: count out of domain
    RETURN;
END_IF

(* 段 3｜空数组恒等：信息级告知后直接成功返回 / Empty array identity: inform and succeed *)
IF nCount = 0 THEN
    uErrorId := 16#0002_303C;    // 信息级：空数组恒等返回 / Info: empty array, identity return
    FC_DL_BytesToHexString := TRUE;
    RETURN;
END_IF

(* 段 4｜逐字节编码：高低半字节各查一次码表 / Encode byte by byte: one table lookup per nibble *)
FOR nI := 0 TO (nCount - 1) DO
    bCur := aBytes[nI];                              // 取当前字节 / Take the current byte
    nHi  := BYTE_TO_INT(SHR(bCur, 4));               // 高半字节 0 到 15 / High nibble, 0 to 15
    nLo  := BYTE_TO_INT(bCur AND 16#0F);             // 低半字节 0 到 15 / Low nibble, 0 to 15
    sTmp := CONCAT(sTmp, MID('0123456789ABCDEF', DL_BTH_ONE, nHi + DL_BTH_ONE)); // 高位字符，下标偏 1 / High char, index shifted
    sTmp := CONCAT(sTmp, MID('0123456789ABCDEF', DL_BTH_ONE, nLo + DL_BTH_ONE)); // 低位字符 / Low char
    nWritten := nWritten + 2;                        // 每字节恒两字符 / Exactly two chars per byte
END_FOR

(* 段 5｜写出一致性校验（防御闸）：长度必须恰为两倍计数 / Consistency gate: length must be twice the count *)
IF (LEN(sTmp) <> nWritten) OR (nWritten <> (2 * nCount)) THEN
    uErrorId := 16#0002_303E;    // 故障级：写出链路异常，结果作废 / Fault: write chain broken, voided
    sHex := '';
    RETURN;
END_IF

(* 段 6｜出口装配：结果与码位单点写出 / Exit: single write for result and code *)
sHex := sTmp;
uErrorId := uCode;
FC_DL_BytesToHexString := TRUE;
END_FUNCTION

(* ---- FC_DL_ByteToBcd.st ---- *)
(*
    FC_DL_ByteToBcd —— 0~99 到 2 位 BCD 的编码
    ------------------------------------------------------------------
    分类      : DL_MathData / Convert
    前缀      : FC_DL_
    版本      : 1.0.0
    溯源      : IEC 61131-3 标准语义的道莅防御性实现（USINT 数值 → BYTE 容器 2 位 BCD）；
                域内委托平台内建 BYTE_TO_BCD，本件不重实现数学内核；
                上域闸门、满量程兜底口径、错误分级与码位 100% 自有；
                clean-room 重写，未复制任何闭源厂商源码，参考实现仅限 MIT/Apache 许可
    平台      : 纯 IEC 61131-3，CODESYS V3.5+ / TwinCAT 3 / InoProShop 通用
    作者      : 道莅代码库 · PLC编程专家（R20）
    ------------------------------------------------------------------
    功能说明  : 把 0~99 的数值编码成 2 位 BCD 写回拨码开关组态字、仪表设定寄存器，
                与 FC_DL_BcdToByte 构成双向对。
                核心防御：① 上域闸门先判：输入 > 99 时不做截断、不做模 100 折算，
                   直接按满量程 16#99 兜底并升故障级——写回方向宁给满量程也不给
                   「半错位值」，因为 100 编码成 16#00 会让设备读到 0，是危险的静默错；
                ② 域内才委托内建，域外调用内建的行为平台间不一致；
                ③ 边界值（0 与 99）发信息级提示，便于排查上游把哨兵值当设定值下发；
                ④ 合成路径（若平台缺内建）按「商 10 / 余 10 拼半字节」落地，
                   域内输入已保证两半字节 ≤ 9，无越界可能。
                职责边界：反向解码归 FC_DL_BcdToByte；4 位 Word 容器归 FC_DL_WordToBcd，
                8 位 Udint 容器归 FC_DL_UdintToBcd；本件只管 2 位拨码容器。
    编译门槛  : 主路径依赖平台内建 BYTE_TO_BCD，三平台标准库均提供。
                若目标平台缺该内建，按合成路径落地：uHi = uIn / 10、uLo = uIn MOD 10
                （两操作数恒为非负且 < 100，取余口径安全），再 uOut = SHL(uHi, 4) OR uLo。
    错误码    : 16#0001_041E 输入恰为域端点（0 或 99），已如实编码——信息级，值可用
                16#0001_041F 预留禁用（信息级，不得挪用）
                16#0001_034B 输入 > 99，已按满量程 16#99 兜底——故障级，bValid = FALSE
                16#0001_034C 预留（故障级，不得挪用）
                16#0001_034D 预留禁用（故障级，不得挪用）
    码位总账  : 16#0001_041E 用 / 16#0001_041F 预留 ｜ 16#0001_034B 用 / 16#0001_034C 预留 / 16#0001_034D 预留
    状态机    : R6 标注 N/A —— 本组件为纯函数无顺序状态机，无 CASE 可写，非法状态不可能出现
    采样约定  : 本件无定时器、无沿检测、无状态；单拍纯计算，结论与任务周期无关。
    修订记录  : 2026-11-16 v1.0.0 首次入库（R20）
*)
FUNCTION FC_DL_ByteToBcd : BYTE
VAR_INPUT
    uIn              : USINT;                 // 输入数值 [无量纲]，有效域 0~99 / input value [dimensionless], valid domain 0 to 99
END_VAR
VAR_OUTPUT
    eErr             : UDINT;                 // 错误码，0=正常 / error id, 0=ok
    bError           : BOOL;                  // 故障标志，eErr 为故障级时 TRUE / error flag, TRUE on fault-level eErr
    bValid           : BOOL;                  // 返回值是否可用（输入越界为 FALSE）/ return usable, FALSE when the input is out of range
END_VAR
VAR CONSTANT
    DL_BCD_IN_MAX    : USINT := 99;           // 2 位 BCD 可表达的数值上限 [无量纲] / the largest value a 2-digit BCD can carry [dimensionless]
    DL_BCD_IN_MIN    : USINT := 0;            // 2 位 BCD 可表达的数值下限 [无量纲] / the smallest value a 2-digit BCD can carry [dimensionless]
    DL_BCD_FULL      : BYTE := 16#99;         // 满量程 BCD 兜底值 [位图] / full scale BCD fallback value [bitmap]
    DL_BYTE_ZERO     : BYTE := 16#00;         // 字节零常量，避免裸字面量 [位图] / byte zero constant [bitmap]
END_VAR
VAR
    uOut             : BYTE;                  // 结果中间量 [位图] / result intermediate [bitmap]
    uWork            : USINT;                 // 入参副本，避免改动调用方数据 [无量纲] / input copy, never modifies caller data [dimensionless]
END_VAR

// 段 1｜返回值与错误状态预置 / segment 1, preset return value and error status
FC_DL_ByteToBcd := DL_BYTE_ZERO;              // 故障缺省返回 0 [位图] / fault default returns zero [bitmap]
eErr := 0;                                    // 预置无错误 / preset no error
bError := FALSE;                              // 预置无故障 / preset no fault
bValid := FALSE;                              // 预置不可用，通过闸门后置位 / preset invalid, set TRUE after the gates
uOut := DL_BYTE_ZERO;                         // 结果中间量清零 / clear the result intermediate
uWork := uIn;                                 // 取入参副本参与判定 / copy the input for the comparisons

// 段 2｜上域闸门：越界即满量程兜底并升故障级（绝不静默截断）/ segment 2, upper gate, full scale fallback with a fault
IF uWork > DL_BCD_IN_MAX THEN
    FC_DL_ByteToBcd := DL_BCD_FULL;           // 满量程兜底 16#99 / fall back to the full scale BCD
    eErr := 16#0001_034B;                     // 故障级：输入超 2 位 BCD 域 / fault level, the input exceeds the 2-digit BCD domain
    bError := TRUE;                           // 置故障标志 / raise the error flag
    bValid := FALSE;                          // 返回值标记不可用 / flag the return as unusable
    RETURN;                                   // 出口，不触碰内建 / exit, the built-in is never touched
END_IF

// 段 3｜主体：域内才委托平台内建 / segment 3, delegate the built-in only inside the domain
uOut := BYTE_TO_BCD(USINT_TO_BYTE(uWork));    // 数值 → BCD 编码 [位图] / encode the number into BCD [bitmap]

// 段 4｜发布结果与域端点提示（信息级，不置 bError）/ segment 4, publish and hint the domain endpoints
FC_DL_ByteToBcd := uOut;                      // 输出 BCD 编码 [位图] / publish the BCD code [bitmap]
bValid := TRUE;                               // 域内编码可用 / the in-domain code is usable
IF (uWork = DL_BCD_IN_MIN) OR (uWork = DL_BCD_IN_MAX) THEN
    eErr := 16#0001_041E;                     // 信息级：输入恰为域端点，多为上游哨兵值 / info level, a domain endpoint, often an upstream sentinel
END_IF
END_FUNCTION

(* ---- FC_DL_CabsComplexCalc.st ---- *)
// FC_DL_CabsComplexCalc v1.0.0
// 开源溯源：brOscatLib / URL https://github.com/iec-oscat-mirror / 许可证 MIT / 借鉴 CABS 复数模长语义（先判大者再缩放，防平方溢出），clean-room 重写
(*
  道莅工业代码库 | DL_MathData | FC_DL_CabsComplexCalc
  版本: 1.0.0 | 日期: 2026-11-23 | 轮次: R75
  功能: 复数模长 |z| = sqrt(re² + im²) 防溢出实现（先判 |re|,|im| 大者，缩放后再平方）
  邻件关系: 与 FC_DL_EuclidDist2DCalc（R74）同防溢出口径族；本件为复数语义命名
            （re/im 实虚部），欧氏件为几何坐标语义（x/y），口径一致不重码
*)
FUNCTION FC_DL_CabsComplexCalc : REAL
VAR_INPUT
    fRe : REAL := 0.0;   // 实部 [无量纲，与虚部同单位] / Real part, same unit as imaginary
    fIm : REAL := 0.0;   // 虚部 [无量纲，与实部同单位] / Imaginary part, same unit as real
END_VAR
VAR_OUTPUT
    bValid : BOOL;       // 结果有效回执 [-] / Result validity receipt
END_VAR
VAR
    fAbsRe : REAL;       // |re| 当拍量 [无量纲] / Absolute real part
    fAbsIm : REAL;       // |im| 当拍量 [无量纲] / Absolute imaginary part
    fMax   : REAL;       // 缩放因子 max(|re|,|im|) [无量纲] / Scaling factor max of both
    fUre   : REAL;       // 缩放后实部 [无量纲] / Scaled real part
    fUim   : REAL;       // 缩放后虚部 [无量纲] / Scaled imaginary part
    fMag   : REAL;       // 缩放域模长 [无量纲] / Magnitude in scaled domain
END_VAR

// —— 段 0：全路径缺省（FC 入口安全侧） —— //
bValid := FALSE;                                   // 有效回执预清 / Validity preset
FC_DL_CabsComplexCalc := 0.0;                      // 返回值缺省安全零 / Return default safe zero

// —— 段 1：非有限闸（NaN 自反判 + 近 Inf 幅值闸） —— //
IF (fRe <> fRe) OR (fIm <> fIm) THEN               // NaN 自反判（判等禁令唯一例外） / NaN self-reflexive test
    RETURN;                                        // 无效返回零 / Invalid, return zero
END_IF
fAbsRe := ABS(fRe);                                // |re| 派生 / Absolute real part
fAbsIm := ABS(fIm);                                // |im| 派生 / Absolute imaginary part
IF (fAbsRe >= 3.0E38) OR (fAbsIm >= 3.0E38) THEN   // 近 Inf 幅值闸（REAL 上限兜底） / Near-Inf magnitude gate
    RETURN;                                        // 无效返回零 / Invalid, return zero
END_IF

// —— 段 2：零向量特判（缩放因子为零时直接归零） —— //
IF (fAbsRe = 0.0) AND (fAbsIm = 0.0) THEN          // 双零特判 / Zero-vector special case
    FC_DL_CabsComplexCalc := 0.0;                  // 模长为零（合法） / Magnitude zero, valid
    bValid := TRUE;                                // 有效回执 / Validity receipt
    RETURN;                                        // 提前返回 / Early return
END_IF

// —— 段 3：防溢出口径（先取大者缩放，再平方求和，杜绝大数平方上溢与小数下溢） —— //
IF fAbsRe >= fAbsIm THEN                           // 取 |re|,|im| 大者为缩放因子 / Larger of the two as factor
    fMax := fAbsRe;
ELSE
    fMax := fAbsIm;
END_IF
fUre := fRe / fMax;                                // 缩放实部 ∈ [-1,1] / Scaled real part in [-1,1]
fUim := fIm / fMax;                                // 缩放虚部 ∈ [-1,1] / Scaled imaginary part in [-1,1]
fMag := SQRT(fUre * fUre + fUim * fUim);           // 缩放域模长 ≤ sqrt(2)，不溢出 / Scaled magnitude <= sqrt(2)
FC_DL_CabsComplexCalc := fMag * fMax;              // 还原真实模长 / Restore true magnitude
bValid := TRUE;                                    // 有效回执 / Validity receipt
END_FUNCTION

(* ---- FC_DL_CalAddMonths.st ---- *)
(*==============================================================================
 * 组件名称 : FC_DL_CalAddMonths ｜ 子库 : DL_MathData ｜ v1.0.0 ｜ 2026-11-24
 * 平台     : CODESYS 3.5 / TwinCAT 3 / InoProShop / Machine Expert（纯 IEC，无厂商库）
 * 功能简介 : 日历加月。给定基准年月日与月增量（可负），输出加月后的年月日，月末钳位：
 *            1 月 31 日 + 1 月 → 2 月 28/29 日；3 月 31 日 − 1 月 → 2 月 28/29 日。
 * 契约     : 合法时返回 TRUE、bValid := TRUE；年/月/日越界（基准日按基准月长度校核）、
 *            |nDelta| > 1200、加月结果落到公元 0 年之前或超出 9999 年 →
 *            返回 FALSE、bError := TRUE、五个出参全部保持 0。
 * 依赖     : 无 DL_ 内部依赖（R16 自足实现：闰年与月长内联），无标准库函数调用
 * 错误码   : R297 零码位范式：eErr 恒 0，仅以 bError / bValid 表达
 * 红线自检 : R1 零全局 R2 零%I/%Q R3 纯IEC R4 除 12 前已证 nIdx 非负且 < 120000
 *            R5 双语注释 R6 N/A（无状态机）R7 N/A（无定时器/沿实例）
 *            R10 仅用 INT_TO_DINT() R11 全声明行分号 R15 标识符零保留字冲突
 * 遗留假设 : 年初口径为公元 1 年 1 月；nDelta 超 ±1200 判故障而非静默截断；
 *            nIdx 为 0 基月序号 = 年 × 12 + 月 − 1 + 增量，非负才可安全除 12 取模。
 * 修订历史 : 2026-11-24 R79-B 首版（日历数论族 1/2）
 *============================================================================*)
FUNCTION FC_DL_CalAddMonths : BOOL
VAR_INPUT
    nYear  : DINT;   // 基准年，公历 1..9999 [年] / base year in the Gregorian range
    nMonth : DINT;   // 基准月，1..12 [月] / base month, one based
    nDay   : DINT;   // 基准日，1..31（按基准月长度校核）[日] / base day checked against the base month length
    nDelta : INT;    // 月增量，可负，|nDelta| ≤ 1200 [月] / month delta, negative allowed
END_VAR
VAR_OUTPUT
    eErr      : UDINT; // 错误码，零码位范式恒 0 / error id, always zero under the zero-code rule
    bError    : BOOL;  // 入参越界或结果不可表示时为真 / TRUE on an input out of range or an unrepresentable result
    bValid    : BOOL;  // 出参可用标志 / TRUE when the outputs are usable
    nOutYear  : DINT;  // 结果年 [年] / resulting year
    nOutMonth : DINT;  // 结果月 1..12 [月] / resulting month
    nOutDay   : DINT;  // 结果日，已按结果月长度钳位 [日] / resulting day clamped to the length of the resulting month
END_VAR
VAR CONSTANT
    DL_ZERO    : DINT := 0;     // 整数零哨兵 / integer zero sentinel
    DL_ONE     : DINT := 1;     // 整数一哨兵 / integer one sentinel
    DL_TWELVE  : DINT := 12;    // 每年月数 [月] / months per year
    DL_D31     : DINT := 31;    // 大月日数上界 [日] / the day count of a long month
    DL_D30     : DINT := 30;    // 小月日数 [日] / the day count of a short month
    DL_D28     : DINT := 28;    // 平年二月日数 [日] / the February day count of a common year
    DL_D29     : DINT := 29;    // 闰年二月日数 [日] / the February day count of a leap year
    DL_YMIN    : DINT := 1;     // 年份下界 [年] / lower year bound
    DL_YMAX    : DINT := 9999;  // 年份上界 [年] / upper year bound
    DL_IDXMAX  : DINT := 120000; // 月序号开区间上界 = 10000 × 12 [月] / exclusive index ceiling
    DL_DMAX    : INT  := 1200;  // 月增量绝对值上界 [月] / absolute month delta ceiling
END_VAR
VAR
    nIdx    : DINT; // 0 基月序号（年 × 12 + 月 − 1 + 增量）[月] / zero based month index
    nMaxDay : DINT; // 基准月的日数 28..31 [日] / days in the base month
    nResMax : DINT; // 结果月的日数 28..31 [日] / days in the resulting month
END_VAR

// 段 1｜出口预置 / segment 1, preset the exit
FC_DL_CalAddMonths := FALSE;  // 缺省失败 / default failure
eErr      := 0;               // 零码位范式 / zero-code rule
bError    := FALSE;           // 预置无故障 / preset no fault
bValid    := FALSE;           // 域闸前不认出参 / the outputs are unusable until the gates pass
nOutYear  := DL_ZERO;         // 年清零 / clear the year
nOutMonth := DL_ZERO;         // 月清零 / clear the month
nOutDay   := DL_ZERO;         // 日清零 / clear the day

// 段 2｜年与月的域闸（含 nDelta 双侧直比，禁 ABS 单侧以免 INT 下界回绕）/ segment 2, the year, month and delta gates
IF (nYear < DL_YMIN) OR (nYear > DL_YMAX) THEN bError := TRUE; RETURN; END_IF              // 年越界 / year out of range
IF (nMonth < DL_ONE) OR (nMonth > DL_TWELVE) THEN bError := TRUE; RETURN; END_IF           // 月越界 / month out of range
IF (nDelta > DL_DMAX) OR (nDelta < -DL_DMAX) THEN bError := TRUE; RETURN; END_IF           // 增量越界 / delta out of range

// 段 3｜基准日校核：按基准月长度，防「2 月 30 日」这类日历不存在日 / segment 3, the base day gate by month length
nMaxDay := DL_D31;                                                                          // 缺省大月 / default to a long month
IF (nMonth = 4) OR (nMonth = 6) OR (nMonth = 9) OR (nMonth = 11) THEN nMaxDay := DL_D30; END_IF  // 小月 / short months
IF nMonth = 2 THEN nMaxDay := DL_D28; END_IF                                               // 二月先按平年 / February as a common year
IF (nMonth = 2) AND (((nYear MOD 4) = 0) AND ((nYear MOD 100) <> 0) OR ((nYear MOD 400) = 0)) THEN nMaxDay := DL_D29; END_IF  // 闰年二月 / leap February
IF (nDay < DL_ONE) OR (nDay > nMaxDay) THEN bError := TRUE; RETURN; END_IF                 // 日越界 / day out of range

// 段 4｜月序号换算与结果域闸（先验后写，出参在故障时保持 0）/ segment 4, the month index and the result domain gate
nIdx := (nYear * DL_TWELVE) + (nMonth - DL_ONE) + INT_TO_DINT(nDelta);                      // 0 基月序号 / the zero based month index
IF (nIdx < DL_ZERO) OR (nIdx >= DL_IDXMAX) THEN bError := TRUE; RETURN; END_IF             // 落到公元 0 年前或超出 9999 年 / before year one or beyond the ceiling
nOutYear  := nIdx / DL_TWELVE;                                                              // 除 12 已证 nIdx 非负 / the division is safe after the non negative gate
nOutMonth := (nIdx MOD DL_TWELVE) + DL_ONE;                                                  // 月序 0..11 加一 / the month index shifted to one based

// 段 5｜月末钳位：结果月短于基准日时收到结果月最后一天 / segment 5, the month end clamp
nResMax := DL_D31;                                                                          // 缺省大月 / default to a long month
IF (nOutMonth = 4) OR (nOutMonth = 6) OR (nOutMonth = 9) OR (nOutMonth = 11) THEN nResMax := DL_D30; END_IF  // 小月 / short months
IF nOutMonth = 2 THEN nResMax := DL_D28; END_IF                                            // 二月先按平年 / February as a common year
IF (nOutMonth = 2) AND (((nOutYear MOD 4) = 0) AND ((nOutYear MOD 100) <> 0) OR ((nOutYear MOD 400) = 0)) THEN nResMax := DL_D29; END_IF  // 闰年二月 / leap February
IF nDay > nResMax THEN nOutDay := nResMax; ELSE nOutDay := nDay; END_IF                     // 钳位 / clamp to the month length
bValid := TRUE;                                                                             // 出参可用 / the outputs are usable
FC_DL_CalAddMonths := TRUE;                                                                 // 加月完成 / the month shift completed
END_FUNCTION

(* ---- FC_DL_CalcDistance2D.st ---- *)
(*
  ==================================================================
  组件名 Component  : FC_DL_CalcDistance2D
  分类   Category   : DL_MathData
  前缀   Naming     : FC_DL_ ｜ b/n/u/f 类型前缀制（R265）
  版本   Version    : 1.0.0
  功能   Purpose    : 2D 平面两点欧氏距离 √(Δx²+Δy²)：大坐标防溢出采用
                      Hypot 等价缩放思路——取 |Δ| 较大者为尺度因子 m，
                      d = m·√((Δx/m)² + (Δy/m)²)，平方项全部落在 1..2，
                      根号项 ≤ √2，杜绝 (1E154)² 型平方溢出。m=0（两点重
                      合）单分支直返 0，不进除法面。
  来源   Source     : t2-1-lgf-math（Hypot 缩放为公开数值方法口径
                      （C99 hypot 语义），实现零源码复制）
  互引   Cross-ref  : FC_DL_CalcDistance3D（同族三维距离件，本件为其平面
                      特例口径属主，二者共用「尺度缩放防溢出」方法论）
  平台   Platform   : 纯 IEC 61131-3 四则 + ABS/SQRT，三平台通用
  依赖   Depends    : 无 DL_ 内部依赖；无标准库
  红线   Redline    : R1 零全局/VAR_EXTERNAL/R2 零 %I/%Q/R3 纯 IEC 标准
                      R4 非有限闸 + 除零闸（m=0 分支）+ 缩放后非有限复核
                      /R5 全变量双语同行注释/R6 纯函数无状态机（CASE 不
                      适用）/R7 无定时器与沿检测/R8 阈值全常量化
  错误码 Codes      : 01【失效级】任一坐标非有限（NaN 自反判 / Inf 上限
                      兜底判），返回 0
                      02【失效级】缩放后中间量或结果非有限（结构性罕见
                      兜底），返回 0
  码位反证 Note     : 01/02 分立依据（R90）：01 在输入面、02 在数值面可
                      观测；02 若并入 01，则「输入全有限仍失败」这一病态
                      信号将不可观测，故必须分立。
  验收   Acceptance : V1 (0,0)-(3,4) → 5 ｜ V2 重合点 → 0（bValid）｜
                      V3 (1E300,0)-(0,1E300) → ≈1.414E300（不溢出）｜
                      V4 含 NaN → 码 01 ｜ V5 两坐标互换 → 距离不变
  变更   Revision   : 2026-11-22  v1.0.0  R67 首版（编码阶段批 2 序 1）
  ==================================================================
*)
FUNCTION FC_DL_CalcDistance2D : LREAL
VAR_INPUT
    fX1    : LREAL;  // 点 1 横坐标 [mm]/[物理单位] / the x of point one
    fY1    : LREAL;  // 点 1 纵坐标 [mm]/[物理单位] / the y of point one
    fX2    : LREAL;  // 点 2 横坐标 [mm]/[物理单位] / the x of point two
    fY2    : LREAL;  // 点 2 纵坐标 [mm]/[物理单位] / the y of point two
END_VAR
VAR_OUTPUT
    bValid : BOOL;   // 距离可用标志 [-] / the distance usable flag
    nErrId : UDINT;  // 错误码，0=正常，01/02 见头注 [码] / the error code [code]
END_VAR
VAR
    fDx    : LREAL;  // 横向增量工作寄存器 / the delta x working register
    fDy    : LREAL;  // 纵向增量工作寄存器 / the delta y working register
    fAx    : LREAL;  // |Δx| 工作寄存器 / the abs delta x register
    fAy    : LREAL;  // |Δy| 工作寄存器 / the abs delta y register
    fScale : LREAL;  // 尺度因子 m = max(|Δx|,|Δy|) / the scale factor m
    fTmp   : LREAL;  // 缩放平方和工作寄存器 / the scaled squared sum register
END_VAR
VAR CONSTANT
    C2D_FIN_MAX  : LREAL := 1.7976931348623157E308; // LREAL 有限上限 / the finite LREAL limit
    C2D_ERR_NONE : UDINT := 16#0000_0000;           // 无错误 [码] / no error [code]
    C2D_ERR_NAN  : UDINT := 16#0000_0001;           // 码 01：输入非有限 / code 01, non finite input
    C2D_ERR_OVF  : UDINT := 16#0000_0002;           // 码 02：中间量/结果非有限 / code 02, non finite intermediate
END_VAR

// 段 1｜输出预置 / segment 1, preset the outputs
FC_DL_CalcDistance2D := 0.0;  // 失效缺省返回 0 / fault default returns zero
bValid := FALSE;              // 预置不可用 / preset unusable
nErrId := C2D_ERR_NONE;       // 预置无错误 / preset no error

// 段 2｜输入非有限闸（码 01）：NaN 自反判 + Inf 上限兜底判 / segment 2, the input finite gate
IF (fX1 <> fX1) OR (fY1 <> fY1) OR (fX2 <> fX2) OR (fY2 <> fY2)
   OR (ABS(fX1) > C2D_FIN_MAX) OR (ABS(fY1) > C2D_FIN_MAX)
   OR (ABS(fX2) > C2D_FIN_MAX) OR (ABS(fY2) > C2D_FIN_MAX) THEN
    nErrId := C2D_ERR_NAN;
    RETURN;
END_IF

// 段 3｜增量与尺度因子（有限值之差仍可能溢出 Inf，段 4 复核）
//      segment 3, the deltas and the scale factor, the finite minus finite can still overflow
fDx := fX2 - fX1;                       // 横向增量 / the delta x
fDy := fY2 - fY1;                       // 纵向增量 / the delta y
fAx := ABS(fDx);                        // |Δx| / the abs delta x
fAy := ABS(fDy);                        // |Δy| / the abs delta y
IF fAx >= fAy THEN                      // 尺度因子取较大者 / the larger magnitude
    fScale := fAx;
ELSE
    fScale := fAy;
END_IF

// 段 4｜重合点分支（m=0 除零闸，直返 0）+ 增量非有限复核（码 01，Inf 归因输入面）
//      segment 4, the coincident point branch and the delta finiteness recheck
IF fScale = 0.0 THEN                    // 两点重合（Δx=Δy=0，零判安全：精确零源自精确相等）/ the coincident points
    FC_DL_CalcDistance2D := 0.0;        // 距离 0 / the zero distance
    bValid := TRUE;                     // 合法零距离 / the valid zero distance
    RETURN;
END_IF
IF (fDx <> fDx) OR (fDy <> fDy) OR (fScale <> fScale) OR (ABS(fDx) > C2D_FIN_MAX) OR (ABS(fDy) > C2D_FIN_MAX) THEN
    nErrId := C2D_ERR_NAN;              // 增量溢出为非有限 / the delta overflowed to non finite
    RETURN;
END_IF

// 段 5｜Hypot 缩放求距：d = m·√((Δx/m)² + (Δy/m)²)，平方项 ∈ 0..1
//      segment 5, the hypot scaled distance, the squared terms inside zero to one
fTmp := (fDx / fScale) * (fDx / fScale) + (fDy / fScale) * (fDy / fScale);  // 缩放平方和 ≤ 2 / the scaled squared sum
IF (fTmp <> fTmp) OR (fTmp < 0.0) OR (fTmp > 2.0000000001) THEN
    nErrId := C2D_ERR_OVF;              // 缩放后仍非有限（结构性罕见兜底）/ the non finite after scaling
    RETURN;
END_IF
FC_DL_CalcDistance2D := fScale * SQRT(fTmp);  // 距离 [mm]/[物理单位] / the distance
IF (FC_DL_CalcDistance2D <> FC_DL_CalcDistance2D) OR (ABS(FC_DL_CalcDistance2D) > C2D_FIN_MAX) THEN
    nErrId := C2D_ERR_OVF;              // 结果非有限复核 / the result finiteness recheck
    FC_DL_CalcDistance2D := 0.0;        // 失效回缺省 0 / fault default zero
    RETURN;
END_IF
bValid := TRUE;                         // 距离可用 / the distance is usable
END_FUNCTION

(* ---- FC_DL_CalDateFromDayOfYear.st ---- *)
(*==============================================================================
 * 组件名称 : FC_DL_CalDateFromDayOfYear ｜ 子库 : DL_MathData ｜ v1.0.1 ｜ 2026-11-24
 * 平台     : CODESYS 3.5 / TwinCAT 3 / InoProShop / Machine Expert（纯 IEC，无厂商库）
 * 功能简介 : 年内序号反解月日 —— 输入公历年与 1~366 的年内序号，出参月、日。
 *            逐月递减法，闰年 2 月按 29 天参与递减。
 * 契约     : 合法时返回 TRUE 并写出 nMonth / nDay；nDayOfYear 越界（<1 或 >当年天数）
 *            或 nYear < 1583 时返回 FALSE、bError := TRUE、nMonth / nDay 均置 0。
 * 依赖     : 无 DL_ 内部依赖（R16 自足实现），无标准库函数调用
 * 错误码   : R297 零码位范式：eErr 恒 0，仅以 bError / bValid 表达
 * 红线自检 : R1 零全局 R2 零%I/%Q R3 纯IEC R4 年份与序号双域闸、无除法
 *            R5 双语注释 R6 N/A（无状态机）R7 N/A（无定时器/沿实例）
 *            R10 无类型转换 R11 全声明行分号 R15 标识符零保留字冲突 R18 N/A（无 bReset）
 * 修订历史 : 2026-11-24 R79-A 首版（日历算术族 4/9）
 *            2026-11-24  v1.0.1  R79/P4：补年份上界闸 DL_GREG_LAST=9999（原仅下界 1583）
 *============================================================================*)
FUNCTION FC_DL_CalDateFromDayOfYear : BOOL
VAR_INPUT
    nYear      : DINT;  // 公历年，域闸 1583 及以上 [年] / Gregorian year, domain starts at 1583 [year]
    nDayOfYear : DINT;  // 年内序号 1~365 或 366 [天] / day of year, one to three hundred sixty six [day]
END_VAR
VAR_OUTPUT
    eErr       : UDINT; // 错误码，零码位范式恒 0 / error id, always zero under the zero-code rule
    bError     : BOOL;  // 序号越界或年份域外为真 / TRUE when the ordinal or the year is out of range
    bValid     : BOOL;  // 出参可用标志 / TRUE when the outputs are usable
    nMonth     : DINT;  // 解出的月份 1~12，故障时 0 [月] / solved month, zero on fault [month]
    nDay       : DINT;  // 解出的日 1~31，故障时 0 [天] / solved day, zero on fault [day]
END_VAR
VAR CONSTANT
    DL_GREG_START : DINT := 1583;   // 格里高利历起点年 [年] / first Gregorian year [year]
    DL_GREG_LAST  : DINT := 9999;   // 年份上界（v1.0.1 补：防 int64/日期串溢出）[年] / Upper year bound added in v1.0.1 [year]
    DL_MONTH_MIN  : DINT := 1;      // 月份下界 [月] / lower month bound [month]
    DL_MONTH_MAX  : DINT := 12;     // 月份上界 [月] / upper month bound [month]
    DL_DAYS_COMMON : DINT := 365;   // 平年天数 [天] / days in a common year [day]
    DL_DAYS_FEB   : DINT := 28;     // 平年 2 月天数 [天] / February days in a common year [day]
    DL_DAYS_30    : DINT := 30;     // 小月天数 [天] / days in a short month [day]
    DL_DAYS_31    : DINT := 31;     // 大月天数 [天] / days in a long month [day]
    DL_STEP4      : DINT := 4;      // 闰年基本步长 [年] / base leap step [year]
    DL_STEP100    : DINT := 100;    // 世纪基数 [年] / century radix [year]
    DL_STEP400    : DINT := 400;    // 四世纪基数 [年] / four century radix [year]
    DL_ZERO       : DINT := 0;      // 整数零哨兵 [无量纲] / integer zero sentinel [dimensionless]
END_VAR
VAR
    bLeap      : BOOL;  // 当年是否闰年 / whether the year is a leap year
    nDaysYear  : DINT;  // 当年总天数 365 或 366 [天] / total days of the year, 365 or 366 [day]
    nRem       : DINT;  // 递减过程中的剩余序号 [天] / remaining ordinal during the walk [day]
    nMonthDays : DINT;  // 当前游标月的天数 [天] / length of the month at the cursor [day]
    i          : DINT;  // 月份游标 1~12 [月] / month cursor from one to twelve [month]
END_VAR

// 段 1｜出口预置 / segment 1, preset the exit
FC_DL_CalDateFromDayOfYear := FALSE;    // 缺省失败 / default failure
eErr     := 0;                          // 零码位范式 / zero-code rule
bError   := FALSE;                      // 预置无故障 / preset no fault
bValid   := FALSE;                      // 域闸前不认出参 / outputs unusable until the gates pass
nMonth   := 0;                          // 月出参清零 / clear the month output
nDay     := 0;                          // 日出参清零 / clear the day output

// 段 2｜域闸：年份 + 年内序号上界（闰年 366） / segment 2, year gate plus the ordinal upper bound
bLeap := (((nYear MOD DL_STEP4) = DL_ZERO) AND ((nYear MOD DL_STEP100) <> DL_ZERO)) OR ((nYear MOD DL_STEP400) = DL_ZERO);
nDaysYear := DL_DAYS_COMMON;
IF bLeap THEN
    nDaysYear := DL_DAYS_COMMON + 1;    // 闰年 366 天 / leap years carry one extra day
END_IF
IF ((nYear < DL_GREG_START) OR (nYear > DL_GREG_LAST)) OR (nDayOfYear < DL_MONTH_MIN) OR (nDayOfYear > nDaysYear) THEN
    bError := TRUE;                     // 年份域外或序号越界 / year out of domain or ordinal out of range
    RETURN;                             // 出参保持 0 / the outputs stay zero
END_IF

// 段 3｜逐月递减：剩余序号超过当月天数即扣减并推进月份 / segment 3, walk the months subtracting their lengths
nRem   := nDayOfYear;                   // 从完整序号起步 / start from the full ordinal
nMonth := DL_MONTH_MIN;                 // 从 1 月起 / start at January
FOR i := DL_MONTH_MIN TO DL_MONTH_MAX DO
    IF i = 2 THEN
        nMonthDays := DL_DAYS_FEB;      // 平年 2 月 / common February
        IF bLeap THEN
            nMonthDays := DL_DAYS_FEB + 1;  // 闰年 2 月 / leap February
        END_IF
    ELSIF (i = 4) OR (i = 6) OR (i = 9) OR (i = 11) THEN
        nMonthDays := DL_DAYS_30;       // 小月 / short month
    ELSE
        nMonthDays := DL_DAYS_31;       // 大月 / long month
    END_IF
    IF nRem > nMonthDays THEN
        nRem   := nRem - nMonthDays;    // 整月扣减 / subtract the whole month
        nMonth := nMonth + 1;           // 月份推进 / advance the month
    END_IF
END_FOR

// 段 4｜出口：剩余序号即日 / segment 4, the leftover ordinal is the day
nDay   := nRem;                         // 1~31 / one to thirty one
bValid := TRUE;                         // 出参可用 / the outputs are usable
FC_DL_CalDateFromDayOfYear := TRUE;     // 转换成功 / conversion succeeded
END_FUNCTION

(* ---- FC_DL_CalDateSpanMonths.st ---- *)
(*==============================================================================
 * 组件名称 : FC_DL_CalDateSpanMonths ｜ 子库 : DL_MathData ｜ v1.0.0 ｜ 2026-11-24
 * 平台     : CODESYS 3.5 / TwinCAT 3 / InoProShop / Machine Expert（纯 IEC，无厂商库）
 * 功能简介 : 两日期之间的整月差（月龄/账龄/保养周期用）。含日修正：月差算出后，
 *            若「结束日 < 起始日」则该月不计（正向再减 1）；反向对称（结束日 > 起始日再加 1）。
 * 契约     : 返回整月差，起始晚于结束返回负值；任一日期非法（年 1..9999、月 1..12、
 *            日超出该月长度）→ 返回 0 并置 bError := TRUE、bValid := FALSE。
 * 依赖     : 无 DL_ 内部依赖（R16 自足实现：闰年与月长内联），无标准库函数调用
 * 错误码   : R297 零码位范式：eErr 恒 0，仅以 bError / bValid 表达
 * 红线自检 : R1 零全局 R2 零%I/%Q R3 纯IEC R4 无除法（只乘 12 与加减）+ 无浮点
 *            R5 双语注释 R6 N/A（无状态机）R7 N/A（无定时器/沿实例）
 *            R10 无类型转换 R11 全声明行分号 R15 标识符零保留字冲突
 * 遗留假设 : 日修正按符号对称，故 Span(a→b) = −Span(b→a) 恒成立；同日不同月按月末口径
 *            计（1 月 31 日 → 2 28 日为 0 个月，非 1 个月）；日修正只看日号不比月长。
 * 修订历史 : 2026-11-24 R79-B 首版（日历数论族 2/2）
 *============================================================================*)
FUNCTION FC_DL_CalDateSpanMonths : DINT
VAR_INPUT
    nYearA  : DINT := 0; // 起始日之年，1..9999 [年] / year of the start date
    nMonthA : DINT := 0; // 起始日之月，1..12 [月] / month of the start date
    nDayA   : DINT := 0; // 起始日之日，1..31 [日] / day of the start date
    nYearB  : DINT := 0; // 结束日之年，1..9999 [年] / year of the end date
    nMonthB : DINT := 0; // 结束日之月，1..12 [月] / month of the end date
    nDayB   : DINT := 0; // 结束日之日，1..31 [日] / day of the end date
END_VAR
VAR_OUTPUT
    eErr   : UDINT; // 错误码，零码位范式恒 0 / error id, always zero under the zero-code rule
    bError : BOOL;  // 任一日期非法时为真 / TRUE when either date is invalid
    bValid : BOOL;  // 返回值可用标志 / TRUE when the return value is usable
END_VAR
VAR CONSTANT
    DL_ZERO   : DINT := 0;     // 整数零哨兵 / integer zero sentinel
    DL_ONE    : DINT := 1;     // 整数一哨兵 / integer one sentinel
    DL_ELEVEN : DINT := 11;    // 小月判定上界之一（11 月）[月] / one of the short month keys
    DL_TWELVE : DINT := 12;    // 每年月数 [月] / months per year
    DL_D31    : DINT := 31;    // 大月日数上界 [日] / the day count of a long month
    DL_D30    : DINT := 30;    // 小月日数 [日] / the day count of a short month
    DL_D28    : DINT := 28;    // 平年二月日数 [日] / the February day count of a common year
    DL_D29    : DINT := 29;    // 闰年二月日数 [日] / the February day count of a leap year
    DL_YMIN   : DINT := 1;     // 年份下界 [年] / lower year bound
    DL_YMAX   : DINT := 9999;  // 年份上界 [年] / upper year bound
END_VAR
VAR
    nMaxA   : DINT; // 起始月的日数 28..31 [日] / days in the start month
    nMaxB   : DINT; // 结束月的日数 28..31 [日] / days in the end month
    nMonths : DINT; // 未做日修正的整月差 [月] / the raw month difference before the day correction
END_VAR

// 段 1｜出口预置 / segment 1, preset the exit
FC_DL_CalDateSpanMonths := DL_ZERO;  // 缺省零 / default zero
eErr   := 0;                          // 零码位范式 / zero-code rule
bError := FALSE;                      // 预置无故障 / preset no fault
bValid := FALSE;                      // 域闸前不认返回值 / the return value is unusable until the gates pass

// 段 2｜两日期的域闸：年/月先行，日按各自月长度（防 2 月 30 日一类不存在日）/ segment 2, the domain gates
IF (nYearA < DL_YMIN) OR (nYearA > DL_YMAX) OR (nYearB < DL_YMIN) OR (nYearB > DL_YMAX) THEN bError := TRUE; RETURN; END_IF      // 年越界 / year out of range
IF (nMonthA < DL_ONE) OR (nMonthA > DL_TWELVE) OR (nMonthB < DL_ONE) OR (nMonthB > DL_TWELVE) THEN bError := TRUE; RETURN; END_IF  // 月越界 / month out of range
nMaxA := DL_D31;                                                                                    // 起始月缺省大月 / start month defaults to long
IF (nMonthA = 4) OR (nMonthA = 6) OR (nMonthA = 9) OR (nMonthA = DL_ELEVEN) THEN nMaxA := DL_D30; END_IF  // 起始小月 / start short month
IF nMonthA = 2 THEN nMaxA := DL_D28; END_IF                                                        // 起始二月按平年 / start February as common year
IF (nMonthA = 2) AND (((nYearA MOD 4) = 0) AND ((nYearA MOD 100) <> 0) OR ((nYearA MOD 400) = 0)) THEN nMaxA := DL_D29; END_IF     // 起始闰二月 / start leap February
nMaxB := DL_D31;                                                                                    // 结束月缺省大月 / end month defaults to long
IF (nMonthB = 4) OR (nMonthB = 6) OR (nMonthB = 9) OR (nMonthB = DL_ELEVEN) THEN nMaxB := DL_D30; END_IF  // 结束小月 / end short month
IF nMonthB = 2 THEN nMaxB := DL_D28; END_IF                                                        // 结束二月按平年 / end February as common year
IF (nMonthB = 2) AND (((nYearB MOD 4) = 0) AND ((nYearB MOD 100) <> 0) OR ((nYearB MOD 400) = 0)) THEN nMaxB := DL_D29; END_IF     // 结束闰二月 / end leap February
IF (nDayA < DL_ONE) OR (nDayA > nMaxA) OR (nDayB < DL_ONE) OR (nDayB > nMaxB) THEN bError := TRUE; RETURN; END_IF                 // 日越界 / day out of range

// 段 3｜未修正整月差：年差乘 12 加月差的代数和（无除法、无溢出风险：年份已限 9999）/ segment 3, the raw month difference
nMonths := ((nYearB - nYearA) * DL_TWELVE) + (nMonthB - nMonthA);                                   // 整月代数和 [月] / signed month difference

// 段 4｜日修正按符号对称分支：正向「结束日 < 起始日」减一，反向「结束日 > 起始日」加一 / segment 4, the sign symmetric day correction
IF nMonths >= DL_ZERO THEN
    IF nDayB < nDayA THEN nMonths := nMonths - DL_ONE; END_IF                                      // 不足以计满一个月 / not a full month yet
ELSE
    IF nDayB > nDayA THEN nMonths := nMonths + DL_ONE; END_IF                                      // 反向对称修正 / the mirrored correction
END_IF

bValid := TRUE;                                    // 返回值可用 / the return value is usable
FC_DL_CalDateSpanMonths := nMonths;                // 回写整月差 / publish the month span
END_FUNCTION

(* ---- FC_DL_CalDayOfYear.st ---- *)
(*==============================================================================
 * 组件名称 : FC_DL_CalDayOfYear ｜ 子库 : DL_MathData ｜ v1.0.1 ｜ 2026-11-24
 * 平台     : CODESYS 3.5 / TwinCAT 3 / InoProShop / Machine Expert（纯 IEC，无厂商库）
 * 功能简介 : 给定公历年月日，返回年内序号 1~366。用儒略日序数相减实现 ——
 *            JDN(年月日) − JDN(同年 1 月 1 日) + 1，闰年自动含入，无需月长表。
 * 契约     : 返回 1~366；nMonth 不在 1~12、nDay 不在当月 1~当月天数、nYear < 1583
 *            时返回 0 且 bError := TRUE。纯函数无状态。
 * 依赖     : 无 DL_ 内部依赖（R16 自足实现），无标准库函数调用
 * 错误码   : R297 零码位范式：eErr 恒 0，仅以 bError / bValid 表达
 * 红线自检 : R1 零全局 R2 零%I/%Q R3 纯IEC R4 域闸三层先行、整数式除数恒正
 *            R5 双语注释 R6 N/A（无状态机）R7 N/A（无定时器/沿实例）
 *            R10 无类型转换 R11 全声明行分号 R15 标识符零保留字冲突 R18 N/A（无 bReset）
 * 遗留假设 : JDN 整数式对 1583 年及以后恒为正，故 1583 为域闸下限；更早年份不入本件。
 * 修订历史 : 2026-11-24 R79-A 首版（日历算术族 3/9）
 *            2026-11-24  v1.0.1  R79/P4：补年份上界闸 DL_GREG_LAST=9999（原仅下界 1583）
 *============================================================================*)
FUNCTION FC_DL_CalDayOfYear : DINT
VAR_INPUT
    nYear     : DINT;   // 公历年，域闸 1583 及以上 [年] / Gregorian year, domain starts at 1583 [year]
    nMonth    : DINT;   // 月份 1~12 [月] / month from one to twelve [month]
    nDay      : DINT;   // 日 1~当月天数 [天] / day from one to the month length [day]
END_VAR
VAR_OUTPUT
    eErr      : UDINT;  // 错误码，零码位范式恒 0 / error id, always zero under the zero-code rule
    bError    : BOOL;   // 日期不存在或域外为真，返回 0 / TRUE when the date is invalid or out of domain, result is zero
    bValid    : BOOL;   // 结果可用标志 / result usable flag
END_VAR
VAR CONSTANT
    DL_GREG_START : DINT := 1583;   // 格里高利历起点年 [年] / first Gregorian year [year]
    DL_GREG_LAST  : DINT := 9999;   // 年份上界（v1.0.1 补：防 int64/日期串溢出）[年] / Upper year bound added in v1.0.1 [year]
    DL_MONTH_MIN  : DINT := 1;      // 月份下界 [月] / lower month bound [month]
    DL_MONTH_MAX  : DINT := 12;     // 月份上界 [月] / upper month bound [month]
    DL_DAYS_FEB   : DINT := 28;     // 平年 2 月天数 [天] / February days in a common year [day]
    DL_DAYS_30    : DINT := 30;     // 小月天数 [天] / days in a short month [day]
    DL_DAYS_31    : DINT := 31;     // 大月天数 [天] / days in a long month [day]
    DL_STEP4      : DINT := 4;      // 闰年基本步长 [年] / base leap step [year]
    DL_STEP100    : DINT := 100;    // 世纪基数 [年] / century radix [year]
    DL_STEP400    : DINT := 400;    // 四世纪基数 [年] / four century radix [year]
    DL_ZERO       : DINT := 0;      // 整数零哨兵 [无量纲] / integer zero sentinel [dimensionless]
END_VAR
VAR
    bLeap      : BOOL;  // 当年是否闰年 / whether the year is a leap year
    nA         : DINT;  // 月份压缩偏置 0 或 1 / month compression offset, zero or one
    nY2        : DINT;  // 儒略式内的世纪内年份 / shifted year inside the Julian formula
    nM2        : DINT;  // 儒略式内的三月基月份 / March based month inside the Julian formula
    nJdn       : DINT;  // 目标日期的儒略日序数 [日] / Julian day number of the requested date [day]
    nJdnJan1   : DINT;  // 同年 1 月 1 日的儒略日序数 [日] / Julian day number of January the first [day]
    nDaysInMon : DINT;  // 当月的实际天数 [天] / actual length of the requested month [day]
END_VAR

// 段 1｜出口预置 / segment 1, preset the exit
FC_DL_CalDayOfYear := 0;        // 缺省 0 / default zero
eErr   := 0;                    // 零码位范式 / zero-code rule
bError := FALSE;                // 预置无故障 / preset no fault
bValid := FALSE;                // 域闸前不认结果 / unusable until the domain gates pass

// 段 2｜域闸：年份 → 月份 → 日，三层依次拦 / segment 2, three domain gates in sequence
IF ((nYear < DL_GREG_START) OR (nYear > DL_GREG_LAST)) OR (nMonth < DL_MONTH_MIN) OR (nMonth > DL_MONTH_MAX) THEN
    bError := TRUE;             // 年份或月份越界 / the year or the month is out of range
    RETURN;                     // 返回 0 / return zero
END_IF
bLeap := (((nYear MOD DL_STEP4) = DL_ZERO) AND ((nYear MOD DL_STEP100) <> DL_ZERO)) OR ((nYear MOD DL_STEP400) = DL_ZERO);
IF nMonth = 2 THEN
    nDaysInMon := DL_DAYS_FEB;      // 平年 2 月 / common February
    IF bLeap THEN
        nDaysInMon := DL_DAYS_FEB + 1;  // 闰年 2 月 / leap February
    END_IF
ELSIF (nMonth = 4) OR (nMonth = 6) OR (nMonth = 9) OR (nMonth = 11) THEN
    nDaysInMon := DL_DAYS_30;       // 小月 / short month
ELSE
    nDaysInMon := DL_DAYS_31;       // 大月 / long month
END_IF
IF (nDay < DL_MONTH_MIN) OR (nDay > nDaysInMon) THEN
    bError := TRUE;             // 日超出当月天数 / the day exceeds the month length
    RETURN;                     // 返回 0 / return zero
END_IF

// 段 3｜儒略日序数：月压缩到三月基，年偏置 4800，偏移 32045 / segment 3, the Julian day number
nA   := (14 - nMonth) / 12;                                  // 1、2 月归上一年的第 13、14 月 / January and February fold into the previous year
nY2  := nYear + 4800 - nA;                                   // 世纪内年份偏置 / shifted year
nM2  := nMonth + 12 * nA - 3;                                // 三月基月份 0~11 / March based month
nJdn := nDay + (153 * nM2 + 2) / 5 + 365 * nY2 + nY2 / DL_STEP4 - nY2 / DL_STEP100 + nY2 / DL_STEP400 - 32045;

// 段 4｜同年 1 月 1 日的序数：m=1、d=1 代入同一式子后化简 / segment 4, ordinal of January the first
nJdnJan1 := 1 + 306 + 365 * (nYear + 4799) + (nYear + 4799) / DL_STEP4 - (nYear + 4799) / DL_STEP100 + (nYear + 4799) / DL_STEP400 - 32045;

// 段 5｜出口：差值加一即年内序号 / segment 5, the difference plus one is the day of year
FC_DL_CalDayOfYear := nJdn - nJdnJan1 + 1;   // 1~366 / one to three hundred sixty six
bValid := TRUE;                              // 日期合法，结果可用 / the date is legal and the result is usable
END_FUNCTION

(* ---- FC_DL_CalIsWeekend.st ---- *)
(*==============================================================================
 * 组件名称 : FC_DL_CalIsWeekend ｜ 子库 : DL_MathData ｜ v1.0.1 ｜ 2026-11-24
 * 平台     : CODESYS 3.5 / TwinCAT 3 / InoProShop / Machine Expert（纯 IEC，无厂商库）
 * 功能简介 : 公历日期是否落在周六或周日。内部以儒略日序数取余得「周一为 0」的星期序号
 *            （JDN MOD 7），序号 ≥ 5 即周末。与 FC_DL_CalWeekdayIndex 同口径但内联
 *            自足实现，不跨件调用（R16）。
 * 契约     : 返回 TRUE=周末；nYear < 1583、nMonth 不在 1~12、nDay 超当月天数时返回 FALSE
 *            且 bValid := FALSE、bError := TRUE（非法日期不得被误判为工作日）。
 * 依赖     : 无 DL_ 内部依赖（R16 自足实现），无标准库函数调用
 * 错误码   : R297 零码位范式：eErr 恒 0，仅以 bError / bValid 表达
 * 红线自检 : R1 零全局 R2 零%I/%Q R3 纯IEC R4 三层域闸先行、取余操作数恒非负
 *            R5 双语注释 R6 N/A（无状态机）R7 N/A（无定时器/沿实例）
 *            R10 无类型转换 R11 全声明行分号 R15 标识符零保留字冲突 R18 N/A（无 bReset）
 * 遗留假设 : 未含法定节假日与调休表 —— 本件只回答「星期几是否落在周末」，
 *            生产排程需另叠节假日日历，不得把本件当班次日历用。
 * 修订历史 : 2026-11-24 R79-A 首版（日历算术族 8/9）
 *            2026-11-24  v1.0.1  R79/P4：补年份上界闸 DL_GREG_LAST=9999（原仅下界 1583）
 *============================================================================*)
FUNCTION FC_DL_CalIsWeekend : BOOL
VAR_INPUT
    nYear     : DINT;   // 公历年，域闸 1583 及以上 [年] / Gregorian year, domain starts at 1583 [year]
    nMonth    : DINT;   // 月份 1~12 [月] / month from one to twelve [month]
    nDay      : DINT;   // 日 1~当月天数 [天] / day from one to the month length [day]
END_VAR
VAR_OUTPUT
    eErr      : UDINT;  // 错误码，零码位范式恒 0 / error id, always zero under the zero-code rule
    bError    : BOOL;   // 日期非法或域外为真 / TRUE when the date is illegal or out of domain
    bValid    : BOOL;   // 结果可用标志 / result usable flag
END_VAR
VAR CONSTANT
    DL_GREG_START : DINT := 1583;   // 格里高利历起点年 [年] / first Gregorian year [year]
    DL_GREG_LAST  : DINT := 9999;   // 年份上界（v1.0.1 补：防 int64/日期串溢出）[年] / Upper year bound added in v1.0.1 [year]
    DL_MONTH_MIN  : DINT := 1;      // 月份与日的下界 [月] / lower bound of the month and the day [month]
    DL_MONTH_MAX  : DINT := 12;     // 月份上界 [月] / upper month bound [month]
    DL_DAYS_FEB   : DINT := 28;     // 平年 2 月天数 [天] / February days in a common year [day]
    DL_DAYS_30    : DINT := 30;     // 小月天数 [天] / days in a short month [day]
    DL_DAYS_31    : DINT := 31;     // 大月天数 [天] / days in a long month [day]
    DL_STEP4      : DINT := 4;      // 闰年基本步长 [年] / base leap step [year]
    DL_STEP100    : DINT := 100;    // 世纪基数 [年] / century radix [year]
    DL_STEP400    : DINT := 400;    // 四世纪基数 [年] / four century radix [year]
    DL_WEEK_MOD   : DINT := 7;      // 星期基数 [天] / weekday radix [day]
    DL_SAT_IDX    : DINT := 5;      // 周一为 0 时周六的序号 / Saturday index when Monday is zero
    DL_ZERO       : DINT := 0;      // 整数零哨兵 [无量纲] / integer zero sentinel [dimensionless]
END_VAR
VAR
    bLeap      : BOOL;  // 当年是否闰年 / whether the year is a leap year
    nDaysInMon : DINT;  // 当月实际天数 [天] / actual length of the month [day]
    nA         : DINT;  // 月份压缩偏置 0 或 1 / month compression offset, zero or one
    nY2        : DINT;  // 儒略式内的世纪内年份 / shifted year inside the Julian formula
    nM2        : DINT;  // 儒略式内的三月基月份 / March based month inside the Julian formula
    nJdn       : DINT;  // 目标日期的儒略日序数 [日] / Julian day number of the requested date [day]
    nDow       : DINT;  // 周一为 0 的星期序号 / weekday index with Monday as zero
END_VAR

// 段 1｜出口预置：缺省非周末 / segment 1, preset the exit to a working day
FC_DL_CalIsWeekend := FALSE;    // 缺省工作日 / default working day
eErr   := 0;                    // 零码位范式 / zero-code rule
bError := FALSE;                // 预置无故障 / preset no fault
bValid := FALSE;                // 域闸前不认结果 / unusable until the domain gates pass

// 段 2｜域闸：年份 → 月份 → 日 / segment 2, three domain gates in sequence
IF ((nYear < DL_GREG_START) OR (nYear > DL_GREG_LAST)) OR (nMonth < DL_MONTH_MIN) OR (nMonth > DL_MONTH_MAX) THEN
    bError := TRUE;             // 年份或月份越界 / the year or the month is out of range
    RETURN;                     // 返回 FALSE / return FALSE
END_IF
bLeap := (((nYear MOD DL_STEP4) = DL_ZERO) AND ((nYear MOD DL_STEP100) <> DL_ZERO)) OR ((nYear MOD DL_STEP400) = DL_ZERO);
IF nMonth = 2 THEN
    nDaysInMon := DL_DAYS_FEB;          // 平年 2 月 / common February
    IF bLeap THEN
        nDaysInMon := DL_DAYS_FEB + 1;  // 闰年 2 月 / leap February
    END_IF
ELSIF (nMonth = 4) OR (nMonth = 6) OR (nMonth = 9) OR (nMonth = 11) THEN
    nDaysInMon := DL_DAYS_30;           // 小月 / short month
ELSE
    nDaysInMon := DL_DAYS_31;           // 大月 / long month
END_IF
IF (nDay < DL_MONTH_MIN) OR (nDay > nDaysInMon) THEN
    bError := TRUE;             // 日超出当月天数 / the day exceeds the month length
    RETURN;                     // 返回 FALSE / return FALSE
END_IF

// 段 3｜儒略日序数与星期序号 / segment 3, the Julian day number and the weekday index
nA   := (14 - nMonth) / 12;                                  // 1、2 月折入上一年 / January and February fold backwards
nY2  := nYear + 4800 - nA;                                   // 世纪内年份偏置 / shifted year
nM2  := nMonth + 12 * nA - 3;                                // 三月基月份 / March based month
nJdn := nDay + (153 * nM2 + 2) / 5 + 365 * nY2 + nY2 / DL_STEP4 - nY2 / DL_STEP100 + nY2 / DL_STEP400 - 32045;
nDow := nJdn MOD DL_WEEK_MOD;                                // 0=周一 … 6=周日 / zero equals Monday

// 段 4｜出口：周六与周日为真 / segment 4, Saturday and Sunday are true
IF nDow >= DL_SAT_IDX THEN
    FC_DL_CalIsWeekend := TRUE;     // 序号 5、6 落在周末 / indexes five and six fall on the weekend
END_IF
bValid := TRUE;                     // 日期合法，结果可用 / the date is legal and the result is usable
END_FUNCTION

(* ---- FC_DL_CalQuarterIndex.st ---- *)
(*==============================================================================
 * 组件名称 : FC_DL_CalQuarterIndex ｜ 子库 : DL_MathData ｜ v1.0.0 ｜ 2026-11-24
 * 平台     : CODESYS 3.5 / TwinCAT 3 / InoProShop / Machine Expert（纯 IEC，无厂商库）
 * 功能简介 : 月份 → 季度序号。整月整除实现：quarter = (month − 1) DIV 3 + 1，
 *            纯整数、无分支表、无浮点。1~3→Q1，4~6→Q2，7~9→Q3，10~12→Q4。
 * 契约     : 返回 1~4；nMonth 不在 1~12 时返回 0、bError := TRUE、bValid := FALSE。
 *            纯函数无状态，同输入同输出，可重入。
 * 依赖     : 无 DL_ 内部依赖（R16 自足实现），无标准库函数调用
 * 错误码   : R297 零码位范式：eErr 恒 0，仅以 bError / bValid 表达
 * 红线自检 : R1 零全局 R2 零%I/%Q R3 纯IEC R4 月份域闸先行、除数恒为常量 3
 *            R5 双语注释 R6 N/A（无状态机）R7 N/A（无定时器/沿实例）
 *            R10 无类型转换 R11 全声明行分号 R15 标识符零保留字冲突 R18 N/A（无 bReset）
 * 修订历史 : 2026-11-24 R79-A 首版（日历算术族 7/9）
 *============================================================================*)
FUNCTION FC_DL_CalQuarterIndex : DINT
VAR_INPUT
    nMonth      : DINT;  // 月份 1~12，越界即故障 [月] / month from one to twelve, out of range is a fault [month]
END_VAR
VAR_OUTPUT
    eErr        : UDINT; // 错误码，零码位范式恒 0 / error id, always zero under the zero-code rule
    bError      : BOOL;  // 月份越界为真 / TRUE when the month is out of range
    bValid      : BOOL;  // 结果可用标志 / result usable flag
END_VAR
VAR CONSTANT
    DL_MONTH_MIN : DINT := 1;   // 月份下界 [月] / lower month bound [month]
    DL_MONTH_MAX : DINT := 12;  // 月份上界 [月] / upper month bound [month]
    DL_MON_PER_Q : DINT := 3;   // 每季度月数 [月] / months per quarter [month]
    DL_Q_MIN     : DINT := 1;   // 季度下界 [季] / lower quarter bound [quarter]
END_VAR

// 段 1｜出口预置 / segment 1, preset the exit
FC_DL_CalQuarterIndex := 0;     // 缺省 0 / default zero
eErr   := 0;                    // 零码位范式 / zero-code rule
bError := FALSE;                // 预置无故障 / preset no fault
bValid := FALSE;                // 域闸前不认结果 / unusable until the domain gate passes

// 段 2｜月份域闸：唯一故障出口 / segment 2, the month domain gate is the only fault exit
IF (nMonth < DL_MONTH_MIN) OR (nMonth > DL_MONTH_MAX) THEN
    bError := TRUE;             // 月份越界 / the month is out of range
    RETURN;                     // 返回 0 / return zero
END_IF

// 段 3｜季度换算：先减一归零基再整除，避免 3、6、9、12 月落到下一季 / segment 3, zero based division
FC_DL_CalQuarterIndex := ((nMonth - DL_MONTH_MIN) / DL_MON_PER_Q) + DL_Q_MIN;   // 1~4 / one to four
bValid := TRUE;                                                                 // 月份入域，结果可用 / the month is legal and the result is usable
END_FUNCTION

(* ---- FC_DL_CeilEx.st ---- *)
(*
    FC_DL_CeilEx —— 向上取整防御包装（向 +∞，DINT 范围钳位 + NaN 拦截）
    ------------------------------------------------------------------
    分类      : DL_MathData / Math-Round
    前缀      : FC_DL_
    版本      : 1.0.0
    溯源      : IEC 61131-3 标准语义的道莅防御性实现
                （内部委托平台内建函数，外围统一错误码/钳位/双语文档；
                  未复制任何闭源厂商源码，参考实现仅限 MIT/Apache 许可）
    平台      : 纯 IEC 61131-3，CODESYS / TwinCAT / InoProShop 通用
    作者      : 道莅代码库 · PLC编程专家（R15）
    ------------------------------------------------------------------
    功能说明  : 向正无穷方向取整（委托内建 CEIL），负小数如 -1.2 得
                -1。NaN 输入拦截返回 0 并置 16#0001_0195；先以 LREAL 承载 CEIL
                结果再做 DINT 范围闸（CEIL 本身不会上溢 LREAL），超
                [-2147483648, 2147483647] 时钳位到边界并置 16#0001_0263，bValid=
                FALSE；无穷输入被范围闸自然拦截。范围内再经 LREAL_TO_DINT
                显式转换，转换永不溢出。
    错误码    : 0000 正常 / 16#0001_0195 入参越界（NaN 已归零） / 16#0001_0263 上溢下溢（已钳位到 DINT 边界）
    修订记录  : 2026-11-16 v1.0.0 首次入库（R15）
*)
FUNCTION FC_DL_CeilEx : DINT
VAR_INPUT
    lrIn : LREAL; // 输入实数 [无量纲]，任意有限值或 NaN/无穷 / input real value [dimensionless], any finite value or NaN/inf
END_VAR
VAR_OUTPUT
    eErr : UDINT; // 错误码，0=正常，1=入参越界，2=上溢下溢 / error id, 0=ok, 1=input out of domain, 2=overflow or underflow
    bError   : BOOL; // 是否出错，eErr 非 0 时为 TRUE / error flag, TRUE when eErr is nonzero
    bValid   : BOOL; // 输出是否有效可用，钳位降级时为 FALSE / output valid, FALSE for clamped degraded results
END_VAR
VAR
    lrR : LREAL; // CEIL 结果中间量 [无量纲]，LREAL 承载不溢出 / intermediate CEIL result [dimensionless], carried in LREAL without overflow
END_VAR
VAR CONSTANT
    DL_CE_HI : LREAL := 2147483647.0; // DINT 上界 [无量纲]，超过即钳位 / DINT upper bound [dimensionless], beyond clamped
    DL_CE_LO : LREAL := -2147483648.0; // DINT 下界 [无量纲]，低于即钳位 / DINT lower bound [dimensionless], below clamped
END_VAR

// 段 1｜返回值与错误状态预置，任何早退路径不留脏码 / segment 1, preset return value and error states
FC_DL_CeilEx := 0; // 返回值预置安全值 0 / preset return to safe value 0
eErr     := 16#0000_0000; // 错误码预置正常 / preset error id to ok
bError       := FALSE; // 错误标志预置无错 / preset error flag to FALSE
bValid       := TRUE; // 有效标志预置可用 / preset valid flag to TRUE

// 段 2｜NaN 拦截：自不等判据，归零早退，不进内核 / segment 2, NaN interception by self-inequality, zeroed early exit
IF lrIn <> lrIn THEN
    eErr := 16#0001_0195; // 信息级：输入 NaN，已归零 / informational, NaN input, zeroed
    bError   := TRUE; // 置错误标志 / raise error flag
    bValid   := FALSE; // 输出不可用 / output invalid
    RETURN; // 返回预置安全值 0 / return preset safe value 0
END_IF

// 段 3｜委托内建 CEIL（向 +∞ 取整），LREAL 承载结果，无穷输入得无穷 / segment 3, delegation to built-in CEIL toward plus infinity, LREAL carry, infinite input stays infinite
lrR := CEIL(lrIn); // 委托内建 CEIL 内核，不自实现取整内核 / delegate to built-in CEIL kernel

// 段 4｜DINT 范围闸：超界钳位并置 16#0001_0263（无穷输入在此被拦截） / segment 4, DINT range gate, clamp beyond bounds with code 2, infinite input intercepted here
IF lrR > DL_CE_HI THEN
    FC_DL_CeilEx := 2147483647; // 上溢钳位到 DINT 上界 / overflow clamped to the DINT upper bound
    eErr     := 16#0001_0263; // 上溢码 / overflow code
    bError       := TRUE; // 置错误标志 / raise error flag
    bValid       := FALSE; // 钳位值非真实取整 / clamped value is not the true ceiling
    RETURN;
ELSIF lrR < DL_CE_LO THEN
    FC_DL_CeilEx := -2147483648; // 下溢钳位到 DINT 下界 / underflow clamped to the DINT lower bound
    eErr     := 16#0001_0263; // 下溢码 / underflow code
    bError       := TRUE; // 置错误标志 / raise error flag
    bValid       := FALSE; // 钳位值非真实取整 / clamped value is not the true ceiling
    RETURN;
END_IF

// 段 5｜范围内显式转换输出（转换永不溢出） / segment 5, explicit in-range conversion and output
FC_DL_CeilEx := LREAL_TO_DINT(lrR); // 范围内显式转换 / explicit in-range conversion
END_FUNCTION

(* ---- FC_DL_CeilToMultipleInt.st ---- *)
(*==============================================================================
 * 组件名称 : FC_DL_CeilToMultipleInt ｜ 子库 : DL_MathData ｜ v1.0.0 ｜ 2026-11-23
 * 平台     : CODESYS 3.5 / TwinCAT 3 / InoProShop / Machine Expert（纯 IEC，无厂商库）
 * 功能简介 : 整数向上（朝 +∞ 方向）对齐到 nMultiple 的倍数。纯整数算术
 *            实现：整除截取得基准，仅当值大于基准时进位一个倍数；
 *            进位前做 DINT 上限反算防饱和溢出，越限饱和到 2147483647。
 * 契约     : 返回向上对齐结果；nMultiple <= 0 恒返回 0；
 *            纯函数无状态、同输入同输出。
 * 依赖     : 无 DL_ 内部依赖（本批自足实现）
 * 红线自检 : R1 零全局 R2 零%I/%Q R3 纯IEC R4 非法倍数返 0 + 上限反算防溢出
 *            R5 双语注释 R6 N/A（无状态机） R7 N/A（无定时器实例）
 * 修订历史 : 2026-11-23 R78-B1 对齐取整族模板派生首版
 *============================================================================*)
FUNCTION FC_DL_CeilToMultipleInt : DINT
VAR_INPUT
    nValue : DINT;          // 输入整数 / Input integer value
    nMultiple : DINT;       // 对齐倍数，须 > 0 / Alignment multiple, must be > 0
END_VAR
VAR
    nLo : DINT;             // 向零截断的基准倍数值 / Truncated-toward-zero base multiple
END_VAR
IF nMultiple <= 0 THEN
    FC_DL_CeilToMultipleInt := 0;       // 非法倍数返 0 / Invalid multiple returns 0
    RETURN;
END_IF
nLo := (nValue / nMultiple) * nMultiple;    // 整除截取得基准 / Base via integer division truncation
IF nValue > nLo THEN
    IF nLo <= (2147483647 - nMultiple) THEN
        nLo := nLo + nMultiple;             // 向 +∞ 对齐到下一倍数 / Align up to next multiple
    ELSE
        nLo := 2147483647;                  // 进位将溢出，饱和到 DINT 上限 / Saturation at DINT max
    END_IF
END_IF
FC_DL_CeilToMultipleInt := nLo;             // 输出向上对齐结果 / Output ceil-aligned result
END_FUNCTION
